(* IEC 61131-3 sources: veristc/veri-stc/tests/st-examples (part 3) *)

cond_a := LimitHigh(raw_070_a, 130);
cond_a := cond_a AND quality_a;
cond_a := cond_a AND (NOT bypass_a);
input_valid_a := InputValid(raw_070_a, 0, 1000);
cond_a := cond_a AND input_valid_a;
IF NOT input_valid_a THEN
    channel_fault_a := channel_fault_a + 1;
END_IF;
cond_b := LimitHigh(raw_070_b, 130);
cond_b := cond_b AND quality_b;
cond_b := cond_b AND (NOT bypass_b);
input_valid_b := InputValid(raw_070_b, 0, 1000);
cond_b := cond_b AND input_valid_b;
IF NOT input_valid_b THEN
    channel_fault_b := channel_fault_b + 1;
END_IF;
cond_c := LimitHigh(raw_070_c, 130);
cond_c := cond_c AND quality_c;
cond_c := cond_c AND (NOT bypass_c);
input_valid_c := InputValid(raw_070_c, 0, 1000);
cond_c := cond_c AND input_valid_c;
IF NOT input_valid_c THEN
    channel_fault_c := channel_fault_c + 1;
END_IF;
cond_d := LimitHigh(raw_070_d, 130);
cond_d := cond_d AND quality_d;
cond_d := cond_d AND (NOT bypass_d);
input_valid_d := InputValid(raw_070_d, 0, 1000);
cond_d := cond_d AND input_valid_d;
IF NOT input_valid_d THEN
    channel_fault_d := channel_fault_d + 1;
END_IF;
vote_ok := TwoOfFour(cond_a, cond_b, cond_c, cond_d);
IF cond_a <> cond_b THEN
    diagnosis_count := diagnosis_count + 1;
END_IF;
IF cond_c <> cond_d THEN
    diagnosis_count := diagnosis_count + 1;
END_IF;
IF NOT vote_ok THEN
    diagnosis_count := diagnosis_count + 1;
END_IF;
latch_a_070 := RS_Next(vote_ok, train_a_reset, latch_a_070);
IF latch_a_070 AND (NOT train_a_inhibit) THEN
    mask_a_08 := mask_a_08 + 64;
    trip_a := 0 < 1;
    scram_a := 0 < 1;
    breaker_a := 0 > 1;
    mfw_a := 0 < 1;
    alarm_a := 0 < 1;
END_IF;
latch_b_070 := RS_Next(vote_ok, train_b_reset, latch_b_070);
IF latch_b_070 AND (NOT train_b_inhibit) THEN
    mask_b_08 := mask_b_08 + 64;
    trip_b := 0 < 1;
    scram_b := 0 < 1;
    breaker_b := 0 > 1;
    mfw_b := 0 < 1;
    alarm_b := 0 < 1;
END_IF;
IF (raw_070_a > 130) AND (NOT cond_a) THEN
    channel_fault_a := channel_fault_a + 1;
END_IF;
IF (raw_070_b > 130) AND (NOT cond_b) THEN
    channel_fault_b := channel_fault_b + 1;
END_IF;
IF (raw_070_c > 130) AND (NOT cond_c) THEN
    channel_fault_c := channel_fault_c + 1;
END_IF;
IF (raw_070_d > 130) AND (NOT cond_d) THEN
    channel_fault_d := channel_fault_d + 1;
END_IF;
IF vote_ok AND train_a_inhibit THEN
    diagnosis_count := diagnosis_count + 1;
END_IF;
IF vote_ok AND train_b_inhibit THEN
    diagnosis_count := diagnosis_count + 1;
END_IF;

cond_a := LimitHigh(raw_071_a, 131);
cond_a := cond_a AND quality_a;
cond_a := cond_a AND (NOT bypass_a);
input_valid_a := InputValid(raw_071_a, 0, 1000);
cond_a := cond_a AND input_valid_a;
IF NOT input_valid_a THEN
    channel_fault_a := channel_fault_a + 1;
END_IF;
cond_b := LimitHigh(raw_071_b, 131);
cond_b := cond_b AND quality_b;
cond_b := cond_b AND (NOT bypass_b);
input_valid_b := InputValid(raw_071_b, 0, 1000);
cond_b := cond_b AND input_valid_b;
IF NOT input_valid_b THEN
    channel_fault_b := channel_fault_b + 1;
END_IF;
cond_c := LimitHigh(raw_071_c, 131);
cond_c := cond_c AND quality_c;
cond_c := cond_c AND (NOT bypass_c);
input_valid_c := InputValid(raw_071_c, 0, 1000);
cond_c := cond_c AND input_valid_c;
IF NOT input_valid_c THEN
    channel_fault_c := channel_fault_c + 1;
END_IF;
cond_d := LimitHigh(raw_071_d, 131);
cond_d := cond_d AND quality_d;
cond_d := cond_d AND (NOT bypass_d);
input_valid_d := InputValid(raw_071_d, 0, 1000);
cond_d := cond_d AND input_valid_d;
IF NOT input_valid_d THEN
    channel_fault_d := channel_fault_d + 1;
END_IF;
vote_ok := TwoOfFour(cond_a, cond_b, cond_c, cond_d);
IF cond_a <> cond_b THEN
    diagnosis_count := diagnosis_count + 1;
END_IF;
IF cond_c <> cond_d THEN
    diagnosis_count := diagnosis_count + 1;
END_IF;
IF NOT vote_ok THEN
    diagnosis_count := diagnosis_count + 1;
END_IF;
latch_a_071 := RS_Next(vote_ok, train_a_reset, latch_a_071);
IF latch_a_071 AND (NOT train_a_inhibit) THEN
    mask_a_08 := mask_a_08 + 128;
    trip_a := 0 < 1;
    scram_a := 0 < 1;
    breaker_a := 0 > 1;
    afw_a := 0 < 1;
    alarm_a := 0 < 1;
END_IF;
latch_b_071 := RS_Next(vote_ok, train_b_reset, latch_b_071);
IF latch_b_071 AND (NOT train_b_inhibit) THEN
    mask_b_08 := mask_b_08 + 128;
    trip_b := 0 < 1;
    scram_b := 0 < 1;
    breaker_b := 0 > 1;
    afw_b := 0 < 1;
    alarm_b := 0 < 1;
END_IF;
IF (raw_071_a > 131) AND (NOT cond_a) THEN
    channel_fault_a := channel_fault_a + 1;
END_IF;
IF (raw_071_b > 131) AND (NOT cond_b) THEN
    channel_fault_b := channel_fault_b + 1;
END_IF;
IF (raw_071_c > 131) AND (NOT cond_c) THEN
    channel_fault_c := channel_fault_c + 1;
END_IF;
IF (raw_071_d > 131) AND (NOT cond_d) THEN
    channel_fault_d := channel_fault_d + 1;
END_IF;
IF vote_ok AND train_a_inhibit THEN
    diagnosis_count := diagnosis_count + 1;
END_IF;
IF vote_ok AND train_b_inhibit THEN
    diagnosis_count := diagnosis_count + 1;
END_IF;

cond_a := LimitHigh(raw_072_a, 132);
cond_a := cond_a AND quality_a;
cond_a := cond_a AND (NOT bypass_a);
input_valid_a := InputValid(raw_072_a, 0, 1000);
cond_a := cond_a AND input_valid_a;
IF NOT input_valid_a THEN
    channel_fault_a := channel_fault_a + 1;
END_IF;
cond_b := LimitHigh(raw_072_b, 132);
cond_b := cond_b AND quality_b;
cond_b := cond_b AND (NOT bypass_b);
input_valid_b := InputValid(raw_072_b, 0, 1000);
cond_b := cond_b AND input_valid_b;
IF NOT input_valid_b THEN
    channel_fault_b := channel_fault_b + 1;
END_IF;
cond_c := LimitHigh(raw_072_c, 132);
cond_c := cond_c AND quality_c;
cond_c := cond_c AND (NOT bypass_c);
input_valid_c := InputValid(raw_072_c, 0, 1000);
cond_c := cond_c AND input_valid_c;
IF NOT input_valid_c THEN
    channel_fault_c := channel_fault_c + 1;
END_IF;
cond_d := LimitHigh(raw_072_d, 132);
cond_d := cond_d AND quality_d;
cond_d := cond_d AND (NOT bypass_d);
input_valid_d := InputValid(raw_072_d, 0, 1000);
cond_d := cond_d AND input_valid_d;
IF NOT input_valid_d THEN
    channel_fault_d := channel_fault_d + 1;
END_IF;
vote_ok := TwoOfFour(cond_a, cond_b, cond_c, cond_d);
IF cond_a <> cond_b THEN
    diagnosis_count := diagnosis_count + 1;
END_IF;
IF cond_c <> cond_d THEN
    diagnosis_count := diagnosis_count + 1;
END_IF;
IF NOT vote_ok THEN
    diagnosis_count := diagnosis_count + 1;
END_IF;
latch_a_072 := RS_Next(vote_ok, train_a_reset, latch_a_072);
IF latch_a_072 AND (NOT train_a_inhibit) THEN
    mask_a_09 := mask_a_09 + 1;
    trip_a := 0 < 1;
    scram_a := 0 < 1;
    breaker_a := 0 > 1;
    si_a := 0 < 1;
    alarm_a := 0 < 1;
END_IF;
latch_b_072 := RS_Next(vote_ok, train_b_reset, latch_b_072);
IF latch_b_072 AND (NOT train_b_inhibit) THEN
    mask_b_09 := mask_b_09 + 1;
    trip_b := 0 < 1;
    scram_b := 0 < 1;
    breaker_b := 0 > 1;
    si_b := 0 < 1;
    alarm_b := 0 < 1;
END_IF;
IF (raw_072_a > 132) AND (NOT cond_a) THEN
    channel_fault_a := channel_fault_a + 1;
END_IF;
IF (raw_072_b > 132) AND (NOT cond_b) THEN
    channel_fault_b := channel_fault_b + 1;
END_IF;
IF (raw_072_c > 132) AND (NOT cond_c) THEN
    channel_fault_c := channel_fault_c + 1;
END_IF;
IF (raw_072_d > 132) AND (NOT cond_d) THEN
    channel_fault_d := channel_fault_d + 1;
END_IF;
IF vote_ok AND train_a_inhibit THEN
    diagnosis_count := diagnosis_count + 1;
END_IF;
IF vote_ok AND train_b_inhibit THEN
    diagnosis_count := diagnosis_count + 1;
END_IF;

cond_a := LimitHigh(raw_073_a, 133);
cond_a := cond_a AND quality_a;
cond_a := cond_a AND (NOT bypass_a);
input_valid_a := InputValid(raw_073_a, 0, 1000);
cond_a := cond_a AND input_valid_a;
IF NOT input_valid_a THEN
    channel_fault_a := channel_fault_a + 1;
END_IF;
cond_b := LimitHigh(raw_073_b, 133);
cond_b := cond_b AND quality_b;
cond_b := cond_b AND (NOT bypass_b);
input_valid_b := InputValid(raw_073_b, 0, 1000);
cond_b := cond_b AND input_valid_b;
IF NOT input_valid_b THEN
    channel_fault_b := channel_fault_b + 1;
END_IF;
cond_c := LimitHigh(raw_073_c, 133);
cond_c := cond_c AND quality_c;
cond_c := cond_c AND (NOT bypass_c);
input_valid_c := InputValid(raw_073_c, 0, 1000);
cond_c := cond_c AND input_valid_c;
IF NOT input_valid_c THEN
    channel_fault_c := channel_fault_c + 1;
END_IF;
cond_d := LimitHigh(raw_073_d, 133);
cond_d := cond_d AND quality_d;
cond_d := cond_d AND (NOT bypass_d);
input_valid_d := InputValid(raw_073_d, 0, 1000);
cond_d := cond_d AND input_valid_d;
IF NOT input_valid_d THEN
    channel_fault_d := channel_fault_d + 1;
END_IF;
vote_ok := TwoOfFour(cond_a, cond_b, cond_c, cond_d);
IF cond_a <> cond_b THEN
    diagnosis_count := diagnosis_count + 1;
END_IF;
IF cond_c <> cond_d THEN
    diagnosis_count := diagnosis_count + 1;
END_IF;
IF NOT vote_ok THEN
    diagnosis_count := diagnosis_count + 1;
END_IF;
latch_a_073 := RS_Next(vote_ok, train_a_reset, latch_a_073);
IF latch_a_073 AND (NOT train_a_inhibit) THEN
    mask_a_09 := mask_a_09 + 2;
    trip_a := 0 < 1;
    scram_a := 0 < 1;
    breaker_a := 0 > 1;
    ci_a := 0 < 1;
    alarm_a := 0 < 1;
END_IF;
latch_b_073 := RS_Next(vote_ok, train_b_reset, latch_b_073);
IF latch_b_073 AND (NOT train_b_inhibit) THEN
    mask_b_09 := mask_b_09 + 2;
    trip_b := 0 < 1;
    scram_b := 0 < 1;
    breaker_b := 0 > 1;
    ci_b := 0 < 1;
    alarm_b := 0 < 1;
END_IF;
IF (raw_073_a > 133) AND (NOT cond_a) THEN
    channel_fault_a := channel_fault_a + 1;
END_IF;
IF (raw_073_b > 133) AND (NOT cond_b) THEN
    channel_fault_b := channel_fault_b + 1;
END_IF;
IF (raw_073_c > 133) AND (NOT cond_c) THEN
    channel_fault_c := channel_fault_c + 1;
END_IF;
IF (raw_073_d > 133) AND (NOT cond_d) THEN
    channel_fault_d := channel_fault_d + 1;
END_IF;
IF vote_ok AND train_a_inhibit THEN
    diagnosis_count := diagnosis_count + 1;
END_IF;
IF vote_ok AND train_b_inhibit THEN
    diagnosis_count := diagnosis_count + 1;
END_IF;

cond_a := LimitHigh(raw_074_a, 134);
cond_a := cond_a AND quality_a;
cond_a := cond_a AND (NOT bypass_a);
input_valid_a := InputValid(raw_074_a, 0, 1000);
cond_a := cond_a AND input_valid_a;
IF NOT input_valid_a THEN
    channel_fault_a := channel_fault_a + 1;
END_IF;
cond_b := LimitHigh(raw_074_b, 134);
cond_b := cond_b AND quality_b;
cond_b := cond_b AND (NOT bypass_b);
input_valid_b := InputValid(raw_074_b, 0, 1000);
cond_b := cond_b AND input_valid_b;
IF NOT input_valid_b THEN
    channel_fault_b := channel_fault_b + 1;
END_IF;
cond_c := LimitHigh(raw_074_c, 134);
cond_c := cond_c AND quality_c;
cond_c := cond_c AND (NOT bypass_c);
input_valid_c := InputValid(raw_074_c, 0, 1000);
cond_c := cond_c AND input_valid_c;
IF NOT input_valid_c THEN
    channel_fault_c := channel_fault_c + 1;
END_IF;
cond_d := LimitHigh(raw_074_d, 134);
cond_d := cond_d AND quality_d;
cond_d := cond_d AND (NOT bypass_d);
input_valid_d := InputValid(raw_074_d, 0, 1000);
cond_d := cond_d AND input_valid_d;
IF NOT input_valid_d THEN
    channel_fault_d := channel_fault_d + 1;
END_IF;
vote_ok := TwoOfFour(cond_a, cond_b, cond_c, cond_d);
IF cond_a <> cond_b THEN
    diagnosis_count := diagnosis_count + 1;
END_IF;
IF cond_c <> cond_d THEN
    diagnosis_count := diagnosis_count + 1;
END_IF;
IF NOT vote_ok THEN
    diagnosis_count := diagnosis_count + 1;
END_IF;
latch_a_074 := RS_Next(vote_ok, train_a_reset, latch_a_074);
IF latch_a_074 AND (NOT train_a_inhibit) THEN
    mask_a_09 := mask_a_09 + 4;
    trip_a := 0 < 1;
    scram_a := 0 < 1;
    breaker_a := 0 > 1;
    mfw_a := 0 < 1;
    alarm_a := 0 < 1;
END_IF;
latch_b_074 := RS_Next(vote_ok, train_b_reset, latch_b_074);
IF latch_b_074 AND (NOT train_b_inhibit) THEN
    mask_b_09 := mask_b_09 + 4;
    trip_b := 0 < 1;
    scram_b := 0 < 1;
    breaker_b := 0 > 1;
    mfw_b := 0 < 1;
    alarm_b := 0 < 1;
END_IF;
IF (raw_074_a > 134) AND (NOT cond_a) THEN
    channel_fault_a := channel_fault_a + 1;
END_IF;
IF (raw_074_b > 134) AND (NOT cond_b) THEN
    channel_fault_b := channel_fault_b + 1;
END_IF;
IF (raw_074_c > 134) AND (NOT cond_c) THEN
    channel_fault_c := channel_fault_c + 1;
END_IF;
IF (raw_074_d > 134) AND (NOT cond_d) THEN
    channel_fault_d := channel_fault_d + 1;
END_IF;
IF vote_ok AND train_a_inhibit THEN
    diagnosis_count := diagnosis_count + 1;
END_IF;
IF vote_ok AND train_b_inhibit THEN
    diagnosis_count := diagnosis_count + 1;
END_IF;

cond_a := LimitHigh(raw_075_a, 135);
cond_a := cond_a AND quality_a;
cond_a := cond_a AND (NOT bypass_a);
input_valid_a := InputValid(raw_075_a, 0, 1000);
cond_a := cond_a AND input_valid_a;
IF NOT input_valid_a THEN
    channel_fault_a := channel_fault_a + 1;
END_IF;
cond_b := LimitHigh(raw_075_b, 135);
cond_b := cond_b AND quality_b;
cond_b := cond_b AND (NOT bypass_b);
input_valid_b := InputValid(raw_075_b, 0, 1000);
cond_b := cond_b AND input_valid_b;
IF NOT input_valid_b THEN
    channel_fault_b := channel_fault_b + 1;
END_IF;
cond_c := LimitHigh(raw_075_c, 135);
cond_c := cond_c AND quality_c;
cond_c := cond_c AND (NOT bypass_c);
input_valid_c := InputValid(raw_075_c, 0, 1000);
cond_c := cond_c AND input_valid_c;
IF NOT input_valid_c THEN
    channel_fault_c := channel_fault_c + 1;
END_IF;
cond_d := LimitHigh(raw_075_d, 135);
cond_d := cond_d AND quality_d;
cond_d := cond_d AND (NOT bypass_d);
input_valid_d := InputValid(raw_075_d, 0, 1000);
cond_d := cond_d AND input_valid_d;
IF NOT input_valid_d THEN
    channel_fault_d := channel_fault_d + 1;
END_IF;
vote_ok := TwoOfFour(cond_a, cond_b, cond_c, cond_d);
IF cond_a <> cond_b THEN
    diagnosis_count := diagnosis_count + 1;
END_IF;
IF cond_c <> cond_d THEN
    diagnosis_count := diagnosis_count + 1;
END_IF;
IF NOT vote_ok THEN
    diagnosis_count := diagnosis_count + 1;
END_IF;
latch_a_075 := RS_Next(vote_ok, train_a_reset, latch_a_075);
IF latch_a_075 AND (NOT train_a_inhibit) THEN
    mask_a_09 := mask_a_09 + 8;
    trip_a := 0 < 1;
    scram_a := 0 < 1;
    breaker_a := 0 > 1;
    afw_a := 0 < 1;
    alarm_a := 0 < 1;
END_IF;
latch_b_075 := RS_Next(vote_ok, train_b_reset, latch_b_075);
IF latch_b_075 AND (NOT train_b_inhibit) THEN
    mask_b_09 := mask_b_09 + 8;
    trip_b := 0 < 1;
    scram_b := 0 < 1;
    breaker_b := 0 > 1;
    afw_b := 0 < 1;
    alarm_b := 0 < 1;
END_IF;
IF (raw_075_a > 135) AND (NOT cond_a) THEN
    channel_fault_a := channel_fault_a + 1;
END_IF;
IF (raw_075_b > 135) AND (NOT cond_b) THEN
    channel_fault_b := channel_fault_b + 1;
END_IF;
IF (raw_075_c > 135) AND (NOT cond_c) THEN
    channel_fault_c := channel_fault_c + 1;
END_IF;
IF (raw_075_d > 135) AND (NOT cond_d) THEN
    channel_fault_d := channel_fault_d + 1;
END_IF;
IF vote_ok AND train_a_inhibit THEN
    diagnosis_count := diagnosis_count + 1;
END_IF;
IF vote_ok AND train_b_inhibit THEN
    diagnosis_count := diagnosis_count + 1;
END_IF;

cond_a := LimitHigh(raw_076_a, 136);
cond_a := cond_a AND quality_a;
cond_a := cond_a AND (NOT bypass_a);
input_valid_a := InputValid(raw_076_a, 0, 1000);
cond_a := cond_a AND input_valid_a;
IF NOT input_valid_a THEN
    channel_fault_a := channel_fault_a + 1;
END_IF;
cond_b := LimitHigh(raw_076_b, 136);
cond_b := cond_b AND quality_b;
cond_b := cond_b AND (NOT bypass_b);
input_valid_b := InputValid(raw_076_b, 0, 1000);
cond_b := cond_b AND input_valid_b;
IF NOT input_valid_b THEN
    channel_fault_b := channel_fault_b + 1;
END_IF;
cond_c := LimitHigh(raw_076_c, 136);
cond_c := cond_c AND quality_c;
cond_c := cond_c AND (NOT bypass_c);
input_valid_c := InputValid(raw_076_c, 0, 1000);
cond_c := cond_c AND input_valid_c;
IF NOT input_valid_c THEN
    channel_fault_c := channel_fault_c + 1;
END_IF;
cond_d := LimitHigh(raw_076_d, 136);
cond_d := cond_d AND quality_d;
cond_d := cond_d AND (NOT bypass_d);
input_valid_d := InputValid(raw_076_d, 0, 1000);
cond_d := cond_d AND input_valid_d;
IF NOT input_valid_d THEN
    channel_fault_d := channel_fault_d + 1;
END_IF;
vote_ok := TwoOfFour(cond_a, cond_b, cond_c, cond_d);
IF cond_a <> cond_b THEN
    diagnosis_count := diagnosis_count + 1;
END_IF;
IF cond_c <> cond_d THEN
    diagnosis_count := diagnosis_count + 1;
END_IF;
IF NOT vote_ok THEN
    diagnosis_count := diagnosis_count + 1;
END_IF;
latch_a_076 := RS_Next(vote_ok, train_a_reset, latch_a_076);
IF latch_a_076 AND (NOT train_a_inhibit) THEN
    mask_a_09 := mask_a_09 + 16;
    trip_a := 0 < 1;
    scram_a := 0 < 1;
    breaker_a := 0 > 1;
    si_a := 0 < 1;
    alarm_a := 0 < 1;
END_IF;
latch_b_076 := RS_Next(vote_ok, train_b_reset, latch_b_076);
IF latch_b_076 AND (NOT train_b_inhibit) THEN
    mask_b_09 := mask_b_09 + 16;
    trip_b := 0 < 1;
    scram_b := 0 < 1;
    breaker_b := 0 > 1;
    si_b := 0 < 1;
    alarm_b := 0 < 1;
END_IF;
IF (raw_076_a > 136) AND (NOT cond_a) THEN
    channel_fault_a := channel_fault_a + 1;
END_IF;
IF (raw_076_b > 136) AND (NOT cond_b) THEN
    channel_fault_b := channel_fault_b + 1;
END_IF;
IF (raw_076_c > 136) AND (NOT cond_c) THEN
    channel_fault_c := channel_fault_c + 1;
END_IF;
IF (raw_076_d > 136) AND (NOT cond_d) THEN
    channel_fault_d := channel_fault_d + 1;
END_IF;
IF vote_ok AND train_a_inhibit THEN
    diagnosis_count := diagnosis_count + 1;
END_IF;
IF vote_ok AND train_b_inhibit THEN
    diagnosis_count := diagnosis_count + 1;
END_IF;

cond_a := LimitHigh(raw_077_a, 137);
cond_a := cond_a AND quality_a;
cond_a := cond_a AND (NOT bypass_a);
input_valid_a := InputValid(raw_077_a, 0, 1000);
cond_a := cond_a AND input_valid_a;
IF NOT input_valid_a THEN
    channel_fault_a := channel_fault_a + 1;
END_IF;
cond_b := LimitHigh(raw_077_b, 137);
cond_b := cond_b AND quality_b;
cond_b := cond_b AND (NOT bypass_b);
input_valid_b := InputValid(raw_077_b, 0, 1000);
cond_b := cond_b AND input_valid_b;
IF NOT input_valid_b THEN
    channel_fault_b := channel_fault_b + 1;
END_IF;
cond_c := LimitHigh(raw_077_c, 137);
cond_c := cond_c AND quality_c;
cond_c := cond_c AND (NOT bypass_c);
input_valid_c := InputValid(raw_077_c, 0, 1000);
cond_c := cond_c AND input_valid_c;
IF NOT input_valid_c THEN
    channel_fault_c := channel_fault_c + 1;
END_IF;
cond_d := LimitHigh(raw_077_d, 137);
cond_d := cond_d AND quality_d;
cond_d := cond_d AND (NOT bypass_d);
input_valid_d := InputValid(raw_077_d, 0, 1000);
cond_d := cond_d AND input_valid_d;
IF NOT input_valid_d THEN
    channel_fault_d := channel_fault_d + 1;
END_IF;
vote_ok := TwoOfFour(cond_a, cond_b, cond_c, cond_d);
IF cond_a <> cond_b THEN
    diagnosis_count := diagnosis_count + 1;
END_IF;
IF cond_c <> cond_d THEN
    diagnosis_count := diagnosis_count + 1;
END_IF;
IF NOT vote_ok THEN
    diagnosis_count := diagnosis_count + 1;
END_IF;
latch_a_077 := RS_Next(vote_ok, train_a_reset, latch_a_077);
IF latch_a_077 AND (NOT train_a_inhibit) THEN
    mask_a_09 := mask_a_09 + 32;
    trip_a := 0 < 1;
    scram_a := 0 < 1;
    breaker_a := 0 > 1;
    ci_a := 0 < 1;
    alarm_a := 0 < 1;
END_IF;
latch_b_077 := RS_Next(vote_ok, train_b_reset, latch_b_077);
IF latch_b_077 AND (NOT train_b_inhibit) THEN
    mask_b_09 := mask_b_09 + 32;
    trip_b := 0 < 1;
    scram_b := 0 < 1;
    breaker_b := 0 > 1;
    ci_b := 0 < 1;
    alarm_b := 0 < 1;
END_IF;
IF (raw_077_a > 137) AND (NOT cond_a) THEN
    channel_fault_a := channel_fault_a + 1;
END_IF;
IF (raw_077_b > 137) AND (NOT cond_b) THEN
    channel_fault_b := channel_fault_b + 1;
END_IF;
IF (raw_077_c > 137) AND (NOT cond_c) THEN
    channel_fault_c := channel_fault_c + 1;
END_IF;
IF (raw_077_d > 137) AND (NOT cond_d) THEN
    channel_fault_d := channel_fault_d + 1;
END_IF;
IF vote_ok AND train_a_inhibit THEN
    diagnosis_count := diagnosis_count + 1;
END_IF;
IF vote_ok AND train_b_inhibit THEN
    diagnosis_count := diagnosis_count + 1;
END_IF;

cond_a := LimitHigh(raw_078_a, 138);
cond_a := cond_a AND quality_a;
cond_a := cond_a AND (NOT bypass_a);
input_valid_a := InputValid(raw_078_a, 0, 1000);
cond_a := cond_a AND input_valid_a;
IF NOT input_valid_a THEN
    channel_fault_a := channel_fault_a + 1;
END_IF;
cond_b := LimitHigh(raw_078_b, 138);
cond_b := cond_b AND quality_b;
cond_b := cond_b AND (NOT bypass_b);
input_valid_b := InputValid(raw_078_b, 0, 1000);
cond_b := cond_b AND input_valid_b;
IF NOT input_valid_b THEN
    channel_fault_b := channel_fault_b + 1;
END_IF;
cond_c := LimitHigh(raw_078_c, 138);
cond_c := cond_c AND quality_c;
cond_c := cond_c AND (NOT bypass_c);
input_valid_c := InputValid(raw_078_c, 0, 1000);
cond_c := cond_c AND input_valid_c;
IF NOT input_valid_c THEN
    channel_fault_c := channel_fault_c + 1;
END_IF;
cond_d := LimitHigh(raw_078_d, 138);
cond_d := cond_d AND quality_d;
cond_d := cond_d AND (NOT bypass_d);
input_valid_d := InputValid(raw_078_d, 0, 1000);
cond_d := cond_d AND input_valid_d;
IF NOT input_valid_d THEN
    channel_fault_d := channel_fault_d + 1;
END_IF;
vote_ok := TwoOfFour(cond_a, cond_b, cond_c, cond_d);
IF cond_a <> cond_b THEN
    diagnosis_count := diagnosis_count + 1;
END_IF;
IF cond_c <> cond_d THEN
    diagnosis_count := diagnosis_count + 1;
END_IF;
IF NOT vote_ok THEN
    diagnosis_count := diagnosis_count + 1;
END_IF;
latch_a_078 := RS_Next(vote_ok, train_a_reset, latch_a_078);
IF latch_a_078 AND (NOT train_a_inhibit) THEN
    mask_a_09 := mask_a_09 + 64;
    trip_a := 0 < 1;
    scram_a := 0 < 1;
    breaker_a := 0 > 1;
    mfw_a := 0 < 1;
    alarm_a := 0 < 1;
END_IF;
latch_b_078 := RS_Next(vote_ok, train_b_reset, latch_b_078);
IF latch_b_078 AND (NOT train_b_inhibit) THEN
    mask_b_09 := mask_b_09 + 64;
    trip_b := 0 < 1;
    scram_b := 0 < 1;
    breaker_b := 0 > 1;
    mfw_b := 0 < 1;
    alarm_b := 0 < 1;
END_IF;
IF (raw_078_a > 138) AND (NOT cond_a) THEN
    channel_fault_a := channel_fault_a + 1;
END_IF;
IF (raw_078_b > 138) AND (NOT cond_b) THEN
    channel_fault_b := channel_fault_b + 1;
END_IF;
IF (raw_078_c > 138) AND (NOT cond_c) THEN
    channel_fault_c := channel_fault_c + 1;
END_IF;
IF (raw_078_d > 138) AND (NOT cond_d) THEN
    channel_fault_d := channel_fault_d + 1;
END_IF;
IF vote_ok AND train_a_inhibit THEN
    diagnosis_count := diagnosis_count + 1;
END_IF;
IF vote_ok AND train_b_inhibit THEN
    diagnosis_count := diagnosis_count + 1;
END_IF;

cond_a := LimitHigh(raw_079_a, 139);
cond_a := cond_a AND quality_a;
cond_a := cond_a AND (NOT bypass_a);
input_valid_a := InputValid(raw_079_a, 0, 1000);
cond_a := cond_a AND input_valid_a;
IF NOT input_valid_a THEN
    channel_fault_a := channel_fault_a + 1;
END_IF;
cond_b := LimitHigh(raw_079_b, 139);
cond_b := cond_b AND quality_b;
cond_b := cond_b AND (NOT bypass_b);
input_valid_b := InputValid(raw_079_b, 0, 1000);
cond_b := cond_b AND input_valid_b;
IF NOT input_valid_b THEN
    channel_fault_b := channel_fault_b + 1;
END_IF;
cond_c := LimitHigh(raw_079_c, 139);
cond_c := cond_c AND quality_c;
cond_c := cond_c AND (NOT bypass_c);
input_valid_c := InputValid(raw_079_c, 0, 1000);
cond_c := cond_c AND input_valid_c;
IF NOT input_valid_c THEN
    channel_fault_c := channel_fault_c + 1;
END_IF;
cond_d := LimitHigh(raw_079_d, 139);
cond_d := cond_d AND quality_d;
cond_d := cond_d AND (NOT bypass_d);
input_valid_d := InputValid(raw_079_d, 0, 1000);
cond_d := cond_d AND input_valid_d;
IF NOT input_valid_d THEN
    channel_fault_d := channel_fault_d + 1;
END_IF;
vote_ok := TwoOfFour(cond_a, cond_b, cond_c, cond_d);
IF cond_a <> cond_b THEN
    diagnosis_count := diagnosis_count + 1;
END_IF;
IF cond_c <> cond_d THEN
    diagnosis_count := diagnosis_count + 1;
END_IF;
IF NOT vote_ok THEN
    diagnosis_count := diagnosis_count + 1;
END_IF;
latch_a_079 := RS_Next(vote_ok, train_a_reset, latch_a_079);
IF latch_a_079 AND (NOT train_a_inhibit) THEN
    mask_a_09 := mask_a_09 + 128;
    trip_a := 0 < 1;
    scram_a := 0 < 1;
    breaker_a := 0 > 1;
    afw_a := 0 < 1;
    alarm_a := 0 < 1;
END_IF;
latch_b_079 := RS_Next(vote_ok, train_b_reset, latch_b_079);
IF latch_b_079 AND (NOT train_b_inhibit) THEN
    mask_b_09 := mask_b_09 + 128;
    trip_b := 0 < 1;
    scram_b := 0 < 1;
    breaker_b := 0 > 1;
    afw_b := 0 < 1;
    alarm_b := 0 < 1;
END_IF;
IF (raw_079_a > 139) AND (NOT cond_a) THEN
    channel_fault_a := channel_fault_a + 1;
END_IF;
IF (raw_079_b > 139) AND (NOT cond_b) THEN
    channel_fault_b := channel_fault_b + 1;
END_IF;
IF (raw_079_c > 139) AND (NOT cond_c) THEN
    channel_fault_c := channel_fault_c + 1;
END_IF;
IF (raw_079_d > 139) AND (NOT cond_d) THEN
    channel_fault_d := channel_fault_d + 1;
END_IF;
IF vote_ok AND train_a_inhibit THEN
    diagnosis_count := diagnosis_count + 1;
END_IF;
IF vote_ok AND train_b_inhibit THEN
    diagnosis_count := diagnosis_count + 1;
END_IF;

cond_a := LimitHigh(raw_080_a, 100);
cond_a := cond_a AND quality_a;
cond_a := cond_a AND (NOT bypass_a);
input_valid_a := InputValid(raw_080_a, 0, 1000);
cond_a := cond_a AND input_valid_a;
IF NOT input_valid_a THEN
    channel_fault_a := channel_fault_a + 1;
END_IF;
cond_b := LimitHigh(raw_080_b, 100);
cond_b := cond_b AND quality_b;
cond_b := cond_b AND (NOT bypass_b);
input_valid_b := InputValid(raw_080_b, 0, 1000);
cond_b := cond_b AND input_valid_b;
IF NOT input_valid_b THEN
    channel_fault_b := channel_fault_b + 1;
END_IF;
cond_c := LimitHigh(raw_080_c, 100);
cond_c := cond_c AND quality_c;
cond_c := cond_c AND (NOT bypass_c);
input_valid_c := InputValid(raw_080_c, 0, 1000);
cond_c := cond_c AND input_valid_c;
IF NOT input_valid_c THEN
    channel_fault_c := channel_fault_c + 1;
END_IF;
cond_d := LimitHigh(raw_080_d, 100);
cond_d := cond_d AND quality_d;
cond_d := cond_d AND (NOT bypass_d);
input_valid_d := InputValid(raw_080_d, 0, 1000);
cond_d := cond_d AND input_valid_d;
IF NOT input_valid_d THEN
    channel_fault_d := channel_fault_d + 1;
END_IF;
vote_ok := TwoOfFour(cond_a, cond_b, cond_c, cond_d);
IF cond_a <> cond_b THEN
    diagnosis_count := diagnosis_count + 1;
END_IF;
IF cond_c <> cond_d THEN
    diagnosis_count := diagnosis_count + 1;
END_IF;
IF NOT vote_ok THEN
    diagnosis_count := diagnosis_count + 1;
END_IF;
latch_a_080 := RS_Next(vote_ok, train_a_reset, latch_a_080);
IF latch_a_080 AND (NOT train_a_inhibit) THEN
    mask_a_10 := mask_a_10 + 1;
    trip_a := 0 < 1;
    scram_a := 0 < 1;
    breaker_a := 0 > 1;
    si_a := 0 < 1;
    alarm_a := 0 < 1;
END_IF;
latch_b_080 := RS_Next(vote_ok, train_b_reset, latch_b_080);
IF latch_b_080 AND (NOT train_b_inhibit) THEN
    mask_b_10 := mask_b_10 + 1;
    trip_b := 0 < 1;
    scram_b := 0 < 1;
    breaker_b := 0 > 1;
    si_b := 0 < 1;
    alarm_b := 0 < 1;
END_IF;
IF (raw_080_a > 100) AND (NOT cond_a) THEN
    channel_fault_a := channel_fault_a + 1;
END_IF;
IF (raw_080_b > 100) AND (NOT cond_b) THEN
    channel_fault_b := channel_fault_b + 1;
END_IF;
IF (raw_080_c > 100) AND (NOT cond_c) THEN
    channel_fault_c := channel_fault_c + 1;
END_IF;
IF (raw_080_d > 100) AND (NOT cond_d) THEN
    channel_fault_d := channel_fault_d + 1;
END_IF;
IF vote_ok AND train_a_inhibit THEN
    diagnosis_count := diagnosis_count + 1;
END_IF;
IF vote_ok AND train_b_inhibit THEN
    diagnosis_count := diagnosis_count + 1;
END_IF;

cond_a := LimitHigh(raw_081_a, 101);
cond_a := cond_a AND quality_a;
cond_a := cond_a AND (NOT bypass_a);
input_valid_a := InputValid(raw_081_a, 0, 1000);
cond_a := cond_a AND input_valid_a;
IF NOT input_valid_a THEN
    channel_fault_a := channel_fault_a + 1;
END_IF;
cond_b := LimitHigh(raw_081_b, 101);
cond_b := cond_b AND quality_b;
cond_b := cond_b AND (NOT bypass_b);
input_valid_b := InputValid(raw_081_b, 0, 1000);
cond_b := cond_b AND input_valid_b;
IF NOT input_valid_b THEN
    channel_fault_b := channel_fault_b + 1;
END_IF;
cond_c := LimitHigh(raw_081_c, 101);
cond_c := cond_c AND quality_c;
cond_c := cond_c AND (NOT bypass_c);
input_valid_c := InputValid(raw_081_c, 0, 1000);
cond_c := cond_c AND input_valid_c;
IF NOT input_valid_c THEN
    channel_fault_c := channel_fault_c + 1;
END_IF;
cond_d := LimitHigh(raw_081_d, 101);
cond_d := cond_d AND quality_d;
cond_d := cond_d AND (NOT bypass_d);
input_valid_d := InputValid(raw_081_d, 0, 1000);
cond_d := cond_d AND input_valid_d;
IF NOT input_valid_d THEN
    channel_fault_d := channel_fault_d + 1;
END_IF;
vote_ok := TwoOfFour(cond_a, cond_b, cond_c, cond_d);
IF cond_a <> cond_b THEN
    diagnosis_count := diagnosis_count + 1;
END_IF;
IF cond_c <> cond_d THEN
    diagnosis_count := diagnosis_count + 1;
END_IF;
IF NOT vote_ok THEN
    diagnosis_count := diagnosis_count + 1;
END_IF;
latch_a_081 := RS_Next(vote_ok, train_a_reset, latch_a_081);
IF latch_a_081 AND (NOT train_a_inhibit) THEN
    mask_a_10 := mask_a_10 + 2;
    trip_a := 0 < 1;
    scram_a := 0 < 1;
    breaker_a := 0 > 1;
    ci_a := 0 < 1;
    alarm_a := 0 < 1;
END_IF;
latch_b_081 := RS_Next(vote_ok, train_b_reset, latch_b_081);
IF latch_b_081 AND (NOT train_b_inhibit) THEN
    mask_b_10 := mask_b_10 + 2;
    trip_b := 0 < 1;
    scram_b := 0 < 1;
    breaker_b := 0 > 1;
    ci_b := 0 < 1;
    alarm_b := 0 < 1;
END_IF;
IF (raw_081_a > 101) AND (NOT cond_a) THEN
    channel_fault_a := channel_fault_a + 1;
END_IF;
IF (raw_081_b > 101) AND (NOT cond_b) THEN
    channel_fault_b := channel_fault_b + 1;
END_IF;
IF (raw_081_c > 101) AND (NOT cond_c) THEN
    channel_fault_c := channel_fault_c + 1;
END_IF;
IF (raw_081_d > 101) AND (NOT cond_d) THEN
    channel_fault_d := channel_fault_d + 1;
END_IF;
IF vote_ok AND train_a_inhibit THEN
    diagnosis_count := diagnosis_count + 1;
END_IF;
IF vote_ok AND train_b_inhibit THEN
    diagnosis_count := diagnosis_count + 1;
END_IF;

cond_a := LimitHigh(raw_082_a, 102);
cond_a := cond_a AND quality_a;
cond_a := cond_a AND (NOT bypass_a);
input_valid_a := InputValid(raw_082_a, 0, 1000);
cond_a := cond_a AND input_valid_a;
IF NOT input_valid_a THEN
    channel_fault_a := channel_fault_a + 1;
END_IF;
cond_b := LimitHigh(raw_082_b, 102);
cond_b := cond_b AND quality_b;
cond_b := cond_b AND (NOT bypass_b);
input_valid_b := InputValid(raw_082_b, 0, 1000);
cond_b := cond_b AND input_valid_b;
IF NOT input_valid_b THEN
    channel_fault_b := channel_fault_b + 1;
END_IF;
cond_c := LimitHigh(raw_082_c, 102);
cond_c := cond_c AND quality_c;
cond_c := cond_c AND (NOT bypass_c);
input_valid_c := InputValid(raw_082_c, 0, 1000);
cond_c := cond_c AND input_valid_c;
IF NOT input_valid_c THEN
    channel_fault_c := channel_fault_c + 1;
END_IF;
cond_d := LimitHigh(raw_082_d, 102);
cond_d := cond_d AND quality_d;
cond_d := cond_d AND (NOT bypass_d);
input_valid_d := InputValid(raw_082_d, 0, 1000);
cond_d := cond_d AND input_valid_d;
IF NOT input_valid_d THEN
    channel_fault_d := channel_fault_d + 1;
END_IF;
vote_ok := TwoOfFour(cond_a, cond_b, cond_c, cond_d);
IF cond_a <> cond_b THEN
    diagnosis_count := diagnosis_count + 1;
END_IF;
IF cond_c <> cond_d THEN
    diagnosis_count := diagnosis_count + 1;
END_IF;
IF NOT vote_ok THEN
    diagnosis_count := diagnosis_count + 1;
END_IF;
latch_a_082 := RS_Next(vote_ok, train_a_reset, latch_a_082);
IF latch_a_082 AND (NOT train_a_inhibit) THEN
    mask_a_10 := mask_a_10 + 4;
    trip_a := 0 < 1;
    scram_a := 0 < 1;
    breaker_a := 0 > 1;
    mfw_a := 0 < 1;
    alarm_a := 0 < 1;
END_IF;
latch_b_082 := RS_Next(vote_ok, train_b_reset, latch_b_082);
IF latch_b_082 AND (NOT train_b_inhibit) THEN
    mask_b_10 := mask_b_10 + 4;
    trip_b := 0 < 1;
    scram_b := 0 < 1;
    breaker_b := 0 > 1;
    mfw_b := 0 < 1;
    alarm_b := 0 < 1;
END_IF;
IF (raw_082_a > 102) AND (NOT cond_a) THEN
    channel_fault_a := channel_fault_a + 1;
END_IF;
IF (raw_082_b > 102) AND (NOT cond_b) THEN
    channel_fault_b := channel_fault_b + 1;
END_IF;
IF (raw_082_c > 102) AND (NOT cond_c) THEN
    channel_fault_c := channel_fault_c + 1;
END_IF;
IF (raw_082_d > 102) AND (NOT cond_d) THEN
    channel_fault_d := channel_fault_d + 1;
END_IF;
IF vote_ok AND train_a_inhibit THEN
    diagnosis_count := diagnosis_count + 1;
END_IF;
IF vote_ok AND train_b_inhibit THEN
    diagnosis_count := diagnosis_count + 1;
END_IF;

cond_a := LimitHigh(raw_083_a, 103);
cond_a := cond_a AND quality_a;
cond_a := cond_a AND (NOT bypass_a);
input_valid_a := InputValid(raw_083_a, 0, 1000);
cond_a := cond_a AND input_valid_a;
IF NOT input_valid_a THEN
    channel_fault_a := channel_fault_a + 1;
END_IF;
cond_b := LimitHigh(raw_083_b, 103);
cond_b := cond_b AND quality_b;
cond_b := cond_b AND (NOT bypass_b);
input_valid_b := InputValid(raw_083_b, 0, 1000);
cond_b := cond_b AND input_valid_b;
IF NOT input_valid_b THEN
    channel_fault_b := channel_fault_b + 1;
END_IF;
cond_c := LimitHigh(raw_083_c, 103);
cond_c := cond_c AND quality_c;
cond_c := cond_c AND (NOT bypass_c);
input_valid_c := InputValid(raw_083_c, 0, 1000);
cond_c := cond_c AND input_valid_c;
IF NOT input_valid_c THEN
    channel_fault_c := channel_fault_c + 1;
END_IF;
cond_d := LimitHigh(raw_083_d, 103);
cond_d := cond_d AND quality_d;
cond_d := cond_d AND (NOT bypass_d);
input_valid_d := InputValid(raw_083_d, 0, 1000);
cond_d := cond_d AND input_valid_d;
IF NOT input_valid_d THEN
    channel_fault_d := channel_fault_d + 1;
END_IF;
vote_ok := TwoOfFour(cond_a, cond_b, cond_c, cond_d);
IF cond_a <> cond_b THEN
    diagnosis_count := diagnosis_count + 1;
END_IF;
IF cond_c <> cond_d THEN
    diagnosis_count := diagnosis_count + 1;
END_IF;
IF NOT vote_ok THEN
    diagnosis_count := diagnosis_count + 1;
END_IF;
latch_a_083 := RS_Next(vote_ok, train_a_reset, latch_a_083);
IF latch_a_083 AND (NOT train_a_inhibit) THEN
    mask_a_10 := mask_a_10 + 8;
    trip_a := 0 < 1;
    scram_a := 0 < 1;
    breaker_a := 0 > 1;
    afw_a := 0 < 1;
    alarm_a := 0 < 1;
END_IF;
latch_b_083 := RS_Next(vote_ok, train_b_reset, latch_b_083);
IF latch_b_083 AND (NOT train_b_inhibit) THEN
    mask_b_10 := mask_b_10 + 8;
    trip_b := 0 < 1;
    scram_b := 0 < 1;
    breaker_b := 0 > 1;
    afw_b := 0 < 1;
    alarm_b := 0 < 1;
END_IF;
IF (raw_083_a > 103) AND (NOT cond_a) THEN
    channel_fault_a := channel_fault_a + 1;
END_IF;
IF (raw_083_b > 103) AND (NOT cond_b) THEN
    channel_fault_b := channel_fault_b + 1;
END_IF;
IF (raw_083_c > 103) AND (NOT cond_c) THEN
    channel_fault_c := channel_fault_c + 1;
END_IF;
IF (raw_083_d > 103) AND (NOT cond_d) THEN
    channel_fault_d := channel_fault_d + 1;
END_IF;
IF vote_ok AND train_a_inhibit THEN
    diagnosis_count := diagnosis_count + 1;
END_IF;
IF vote_ok AND train_b_inhibit THEN
    diagnosis_count := diagnosis_count + 1;
END_IF;

cond_a := LimitHigh(raw_084_a, 104);
cond_a := cond_a AND quality_a;
cond_a := cond_a AND (NOT bypass_a);
input_valid_a := InputValid(raw_084_a, 0, 1000);
cond_a := cond_a AND input_valid_a;
IF NOT input_valid_a THEN
    channel_fault_a := channel_fault_a + 1;
END_IF;
cond_b := LimitHigh(raw_084_b, 104);
cond_b := cond_b AND quality_b;
cond_b := cond_b AND (NOT bypass_b);
input_valid_b := InputValid(raw_084_b, 0, 1000);
cond_b := cond_b AND input_valid_b;
IF NOT input_valid_b THEN
    channel_fault_b := channel_fault_b + 1;
END_IF;
cond_c := LimitHigh(raw_084_c, 104);
cond_c := cond_c AND quality_c;
cond_c := cond_c AND (NOT bypass_c);
input_valid_c := InputValid(raw_084_c, 0, 1000);
cond_c := cond_c AND input_valid_c;
IF NOT input_valid_c THEN
    channel_fault_c := channel_fault_c + 1;
END_IF;
cond_d := LimitHigh(raw_084_d, 104);
cond_d := cond_d AND quality_d;
cond_d := cond_d AND (NOT bypass_d);
input_valid_d := InputValid(raw_084_d, 0, 1000);
cond_d := cond_d AND input_valid_d;
IF NOT input_valid_d THEN
    channel_fault_d := channel_fault_d + 1;
END_IF;
vote_ok := TwoOfFour(cond_a, cond_b, cond_c, cond_d);
IF cond_a <> cond_b THEN
    diagnosis_count := diagnosis_count + 1;
END_IF;
IF cond_c <> cond_d THEN
    diagnosis_count := diagnosis_count + 1;
END_IF;
IF NOT vote_ok THEN
    diagnosis_count := diagnosis_count + 1;
END_IF;
latch_a_084 := RS_Next(vote_ok, train_a_reset, latch_a_084);
IF latch_a_084 AND (NOT train_a_inhibit) THEN
    mask_a_10 := mask_a_10 + 16;
    trip_a := 0 < 1;
    scram_a := 0 < 1;
    breaker_a := 0 > 1;
    si_a := 0 < 1;
    alarm_a := 0 < 1;
END_IF;
latch_b_084 := RS_Next(vote_ok, train_b_reset, latch_b_084);
IF latch_b_084 AND (NOT train_b_inhibit) THEN
    mask_b_10 := mask_b_10 + 16;
    trip_b := 0 < 1;
    scram_b := 0 < 1;
    breaker_b := 0 > 1;
    si_b := 0 < 1;
    alarm_b := 0 < 1;
END_IF;
IF (raw_084_a > 104) AND (NOT cond_a) THEN
    channel_fault_a := channel_fault_a + 1;
END_IF;
IF (raw_084_b > 104) AND (NOT cond_b) THEN
    channel_fault_b := channel_fault_b + 1;
END_IF;
IF (raw_084_c > 104) AND (NOT cond_c) THEN
    channel_fault_c := channel_fault_c + 1;
END_IF;
IF (raw_084_d > 104) AND (NOT cond_d) THEN
    channel_fault_d := channel_fault_d + 1;
END_IF;
IF vote_ok AND train_a_inhibit THEN
    diagnosis_count := diagnosis_count + 1;
END_IF;
IF vote_ok AND train_b_inhibit THEN
    diagnosis_count := diagnosis_count + 1;
END_IF;

cond_a := LimitHigh(raw_085_a, 105);
cond_a := cond_a AND quality_a;
cond_a := cond_a AND (NOT bypass_a);
input_valid_a := InputValid(raw_085_a, 0, 1000);
cond_a := cond_a AND input_valid_a;
IF NOT input_valid_a THEN
    channel_fault_a := channel_fault_a + 1;
END_IF;
cond_b := LimitHigh(raw_085_b, 105);
cond_b := cond_b AND quality_b;
cond_b := cond_b AND (NOT bypass_b);
input_valid_b := InputValid(raw_085_b, 0, 1000);
cond_b := cond_b AND input_valid_b;
IF NOT input_valid_b THEN
    channel_fault_b := channel_fault_b + 1;
END_IF;
cond_c := LimitHigh(raw_085_c, 105);
cond_c := cond_c AND quality_c;
cond_c := cond_c AND (NOT bypass_c);
input_valid_c := InputValid(raw_085_c, 0, 1000);
cond_c := cond_c AND input_valid_c;
IF NOT input_valid_c THEN
    channel_fault_c := channel_fault_c + 1;
END_IF;
cond_d := LimitHigh(raw_085_d, 105);
cond_d := cond_d AND quality_d;
cond_d := cond_d AND (NOT bypass_d);
input_valid_d := InputValid(raw_085_d, 0, 1000);
cond_d := cond_d AND input_valid_d;
IF NOT input_valid_d THEN
    channel_fault_d := channel_fault_d + 1;
END_IF;
vote_ok := TwoOfFour(cond_a, cond_b, cond_c, cond_d);
IF cond_a <> cond_b THEN
    diagnosis_count := diagnosis_count + 1;
END_IF;
IF cond_c <> cond_d THEN
    diagnosis_count := diagnosis_count + 1;
END_IF;
IF NOT vote_ok THEN
    diagnosis_count := diagnosis_count + 1;
END_IF;
latch_a_085 := RS_Next(vote_ok, train_a_reset, latch_a_085);
IF latch_a_085 AND (NOT train_a_inhibit) THEN
    mask_a_10 := mask_a_10 + 32;
    trip_a := 0 < 1;
    scram_a := 0 < 1;
    breaker_a := 0 > 1;
    ci_a := 0 < 1;
    alarm_a := 0 < 1;
END_IF;
latch_b_085 := RS_Next(vote_ok, train_b_reset, latch_b_085);
IF latch_b_085 AND (NOT train_b_inhibit) THEN
    mask_b_10 := mask_b_10 + 32;
    trip_b := 0 < 1;
    scram_b := 0 < 1;
    breaker_b := 0 > 1;
    ci_b := 0 < 1;
    alarm_b := 0 < 1;
END_IF;
IF (raw_085_a > 105) AND (NOT cond_a) THEN
    channel_fault_a := channel_fault_a + 1;
END_IF;
IF (raw_085_b > 105) AND (NOT cond_b) THEN
    channel_fault_b := channel_fault_b + 1;
END_IF;
IF (raw_085_c > 105) AND (NOT cond_c) THEN
    channel_fault_c := channel_fault_c + 1;
END_IF;
IF (raw_085_d > 105) AND (NOT cond_d) THEN
    channel_fault_d := channel_fault_d + 1;
END_IF;
IF vote_ok AND train_a_inhibit THEN
    diagnosis_count := diagnosis_count + 1;
END_IF;
IF vote_ok AND train_b_inhibit THEN
    diagnosis_count := diagnosis_count + 1;
END_IF;

cond_a := LimitHigh(raw_086_a, 106);
cond_a := cond_a AND quality_a;
cond_a := cond_a AND (NOT bypass_a);
input_valid_a := InputValid(raw_086_a, 0, 1000);
cond_a := cond_a AND input_valid_a;
IF NOT input_valid_a THEN
    channel_fault_a := channel_fault_a + 1;
END_IF;
cond_b := LimitHigh(raw_086_b, 106);
cond_b := cond_b AND quality_b;
cond_b := cond_b AND (NOT bypass_b);
input_valid_b := InputValid(raw_086_b, 0, 1000);
cond_b := cond_b AND input_valid_b;
IF NOT input_valid_b THEN
    channel_fault_b := channel_fault_b + 1;
END_IF;
cond_c := LimitHigh(raw_086_c, 106);
cond_c := cond_c AND quality_c;
cond_c := cond_c AND (NOT bypass_c);
input_valid_c := InputValid(raw_086_c, 0, 1000);
cond_c := cond_c AND input_valid_c;
IF NOT input_valid_c THEN
    channel_fault_c := channel_fault_c + 1;
END_IF;
cond_d := LimitHigh(raw_086_d, 106);
cond_d := cond_d AND quality_d;
cond_d := cond_d AND (NOT bypass_d);
input_valid_d := InputValid(raw_086_d, 0, 1000);
cond_d := cond_d AND input_valid_d;
IF NOT input_valid_d THEN
    channel_fault_d := channel_fault_d + 1;
END_IF;
vote_ok := TwoOfFour(cond_a, cond_b, cond_c, cond_d);
IF cond_a <> cond_b THEN
    diagnosis_count := diagnosis_count + 1;
END_IF;
IF cond_c <> cond_d THEN
    diagnosis_count := diagnosis_count + 1;
END_IF;
IF NOT vote_ok THEN
    diagnosis_count := diagnosis_count + 1;
END_IF;
latch_a_086 := RS_Next(vote_ok, train_a_reset, latch_a_086);
IF latch_a_086 AND (NOT train_a_inhibit) THEN
    mask_a_10 := mask_a_10 + 64;
    trip_a := 0 < 1;
    scram_a := 0 < 1;
    breaker_a := 0 > 1;
    mfw_a := 0 < 1;
    alarm_a := 0 < 1;
END_IF;
latch_b_086 := RS_Next(vote_ok, train_b_reset, latch_b_086);
IF latch_b_086 AND (NOT train_b_inhibit) THEN
    mask_b_10 := mask_b_10 + 64;
    trip_b := 0 < 1;
    scram_b := 0 < 1;
    breaker_b := 0 > 1;
    mfw_b := 0 < 1;
    alarm_b := 0 < 1;
END_IF;
IF (raw_086_a > 106) AND (NOT cond_a) THEN
    channel_fault_a := channel_fault_a + 1;
END_IF;
IF (raw_086_b > 106) AND (NOT cond_b) THEN
    channel_fault_b := channel_fault_b + 1;
END_IF;
IF (raw_086_c > 106) AND (NOT cond_c) THEN
    channel_fault_c := channel_fault_c + 1;
END_IF;
IF (raw_086_d > 106) AND (NOT cond_d) THEN
    channel_fault_d := channel_fault_d + 1;
END_IF;
IF vote_ok AND train_a_inhibit THEN
    diagnosis_count := diagnosis_count + 1;
END_IF;
IF vote_ok AND train_b_inhibit THEN
    diagnosis_count := diagnosis_count + 1;
END_IF;

cond_a := LimitHigh(raw_087_a, 107);
cond_a := cond_a AND quality_a;
cond_a := cond_a AND (NOT bypass_a);
input_valid_a := InputValid(raw_087_a, 0, 1000);
cond_a := cond_a AND input_valid_a;
IF NOT input_valid_a THEN
    channel_fault_a := channel_fault_a + 1;
END_IF;
cond_b := LimitHigh(raw_087_b, 107);
cond_b := cond_b AND quality_b;
cond_b := cond_b AND (NOT bypass_b);
input_valid_b := InputValid(raw_087_b, 0, 1000);
cond_b := cond_b AND input_valid_b;
IF NOT input_valid_b THEN
    channel_fault_b := channel_fault_b + 1;
END_IF;
cond_c := LimitHigh(raw_087_c, 107);
cond_c := cond_c AND quality_c;
cond_c := cond_c AND (NOT bypass_c);
input_valid_c := InputValid(raw_087_c, 0, 1000);
cond_c := cond_c AND input_valid_c;
IF NOT input_valid_c THEN
    channel_fault_c := channel_fault_c + 1;
END_IF;
cond_d := LimitHigh(raw_087_d, 107);
cond_d := cond_d AND quality_d;
cond_d := cond_d AND (NOT bypass_d);
input_valid_d := InputValid(raw_087_d, 0, 1000);
cond_d := cond_d AND input_valid_d;
IF NOT input_valid_d THEN
    channel_fault_d := channel_fault_d + 1;
END_IF;
vote_ok := TwoOfFour(cond_a, cond_b, cond_c, cond_d);
IF cond_a <> cond_b THEN
    diagnosis_count := diagnosis_count + 1;
END_IF;
IF cond_c <> cond_d THEN
    diagnosis_count := diagnosis_count + 1;
END_IF;
IF NOT vote_ok THEN
    diagnosis_count := diagnosis_count + 1;
END_IF;
latch_a_087 := RS_Next(vote_ok, train_a_reset, latch_a_087);
IF latch_a_087 AND (NOT train_a_inhibit) THEN
    mask_a_10 := mask_a_10 + 128;
    trip_a := 0 < 1;
    scram_a := 0 < 1;
    breaker_a := 0 > 1;
    afw_a := 0 < 1;
    alarm_a := 0 < 1;
END_IF;
latch_b_087 := RS_Next(vote_ok, train_b_reset, latch_b_087);
IF latch_b_087 AND (NOT train_b_inhibit) THEN
    mask_b_10 := mask_b_10 + 128;
    trip_b := 0 < 1;
    scram_b := 0 < 1;
    breaker_b := 0 > 1;
    afw_b := 0 < 1;
    alarm_b := 0 < 1;
END_IF;
IF (raw_087_a > 107) AND (NOT cond_a) THEN
    channel_fault_a := channel_fault_a + 1;
END_IF;
IF (raw_087_b > 107) AND (NOT cond_b) THEN
    channel_fault_b := channel_fault_b + 1;
END_IF;
IF (raw_087_c > 107) AND (NOT cond_c) THEN
    channel_fault_c := channel_fault_c + 1;
END_IF;
IF (raw_087_d > 107) AND (NOT cond_d) THEN
    channel_fault_d := channel_fault_d + 1;
END_IF;
IF vote_ok AND train_a_inhibit THEN
    diagnosis_count := diagnosis_count + 1;
END_IF;
IF vote_ok AND train_b_inhibit THEN
    diagnosis_count := diagnosis_count + 1;
END_IF;

cond_a := LimitHigh(raw_088_a, 108);
cond_a := cond_a AND quality_a;
cond_a := cond_a AND (NOT bypass_a);
input_valid_a := InputValid(raw_088_a, 0, 1000);
cond_a := cond_a AND input_valid_a;
IF NOT input_valid_a THEN
    channel_fault_a := channel_fault_a + 1;
END_IF;
cond_b := LimitHigh(raw_088_b, 108);
cond_b := cond_b AND quality_b;
cond_b := cond_b AND (NOT bypass_b);
input_valid_b := InputValid(raw_088_b, 0, 1000);
cond_b := cond_b AND input_valid_b;
IF NOT input_valid_b THEN
    channel_fault_b := channel_fault_b + 1;
END_IF;
cond_c := LimitHigh(raw_088_c, 108);
cond_c := cond_c AND quality_c;
cond_c := cond_c AND (NOT bypass_c);
input_valid_c := InputValid(raw_088_c, 0, 1000);
cond_c := cond_c AND input_valid_c;
IF NOT input_valid_c THEN
    channel_fault_c := channel_fault_c + 1;
END_IF;
cond_d := LimitHigh(raw_088_d, 108);
cond_d := cond_d AND quality_d;
cond_d := cond_d AND (NOT bypass_d);
input_valid_d := InputValid(raw_088_d, 0, 1000);
cond_d := cond_d AND input_valid_d;
IF NOT input_valid_d THEN
    channel_fault_d := channel_fault_d + 1;
END_IF;
vote_ok := TwoOfFour(cond_a, cond_b, cond_c, cond_d);
IF cond_a <> cond_b THEN
    diagnosis_count := diagnosis_count + 1;
END_IF;
IF cond_c <> cond_d THEN
    diagnosis_count := diagnosis_count + 1;
END_IF;
IF NOT vote_ok THEN
    diagnosis_count := diagnosis_count + 1;
END_IF;
latch_a_088 := RS_Next(vote_ok, train_a_reset, latch_a_088);
IF latch_a_088 AND (NOT train_a_inhibit) THEN
    mask_a_11 := mask_a_11 + 1;
    trip_a := 0 < 1;
    scram_a := 0 < 1;
    breaker_a := 0 > 1;
    si_a := 0 < 1;
    alarm_a := 0 < 1;
END_IF;
latch_b_088 := RS_Next(vote_ok, train_b_reset, latch_b_088);
IF latch_b_088 AND (NOT train_b_inhibit) THEN
    mask_b_11 := mask_b_11 + 1;
    trip_b := 0 < 1;
    scram_b := 0 < 1;
    breaker_b := 0 > 1;
    si_b := 0 < 1;
    alarm_b := 0 < 1;
END_IF;
IF (raw_088_a > 108) AND (NOT cond_a) THEN
    channel_fault_a := channel_fault_a + 1;
END_IF;
IF (raw_088_b > 108) AND (NOT cond_b) THEN
    channel_fault_b := channel_fault_b + 1;
END_IF;
IF (raw_088_c > 108) AND (NOT cond_c) THEN
    channel_fault_c := channel_fault_c + 1;
END_IF;
IF (raw_088_d > 108) AND (NOT cond_d) THEN
    channel_fault_d := channel_fault_d + 1;
END_IF;
IF vote_ok AND train_a_inhibit THEN
    diagnosis_count := diagnosis_count + 1;
END_IF;
IF vote_ok AND train_b_inhibit THEN
    diagnosis_count := diagnosis_count + 1;
END_IF;

cond_a := LimitHigh(raw_089_a, 109);
cond_a := cond_a AND quality_a;
cond_a := cond_a AND (NOT bypass_a);
input_valid_a := InputValid(raw_089_a, 0, 1000);
cond_a := cond_a AND input_valid_a;
IF NOT input_valid_a THEN
    channel_fault_a := channel_fault_a + 1;
END_IF;
cond_b := LimitHigh(raw_089_b, 109);
cond_b := cond_b AND quality_b;
cond_b := cond_b AND (NOT bypass_b);
input_valid_b := InputValid(raw_089_b, 0, 1000);
cond_b := cond_b AND input_valid_b;
IF NOT input_valid_b THEN
    channel_fault_b := channel_fault_b + 1;
END_IF;
cond_c := LimitHigh(raw_089_c, 109);
cond_c := cond_c AND quality_c;
cond_c := cond_c AND (NOT bypass_c);
input_valid_c := InputValid(raw_089_c, 0, 1000);
cond_c := cond_c AND input_valid_c;
IF NOT input_valid_c THEN
    channel_fault_c := channel_fault_c + 1;
END_IF;
cond_d := LimitHigh(raw_089_d, 109);
cond_d := cond_d AND quality_d;
cond_d := cond_d AND (NOT bypass_d);
input_valid_d := InputValid(raw_089_d, 0, 1000);
cond_d := cond_d AND input_valid_d;
IF NOT input_valid_d THEN
    channel_fault_d := channel_fault_d + 1;
END_IF;
vote_ok := TwoOfFour(cond_a, cond_b, cond_c, cond_d);
IF cond_a <> cond_b THEN
    diagnosis_count := diagnosis_count + 1;
END_IF;
IF cond_c <> cond_d THEN
    diagnosis_count := diagnosis_count + 1;
END_IF;
IF NOT vote_ok THEN
    diagnosis_count := diagnosis_count + 1;
END_IF;
latch_a_089 := RS_Next(vote_ok, train_a_reset, latch_a_089);
IF latch_a_089 AND (NOT train_a_inhibit) THEN
    mask_a_11 := mask_a_11 + 2;
    trip_a := 0 < 1;
    scram_a := 0 < 1;
    breaker_a := 0 > 1;
    ci_a := 0 < 1;
    alarm_a := 0 < 1;
END_IF;
latch_b_089 := RS_Next(vote_ok, train_b_reset, latch_b_089);
IF latch_b_089 AND (NOT train_b_inhibit) THEN
    mask_b_11 := mask_b_11 + 2;
    trip_b := 0 < 1;
    scram_b := 0 < 1;
    breaker_b := 0 > 1;
    ci_b := 0 < 1;
    alarm_b := 0 < 1;
END_IF;
IF (raw_089_a > 109) AND (NOT cond_a) THEN
    channel_fault_a := channel_fault_a + 1;
END_IF;
IF (raw_089_b > 109) AND (NOT cond_b) THEN
    channel_fault_b := channel_fault_b + 1;
END_IF;
IF (raw_089_c > 109) AND (NOT cond_c) THEN
    channel_fault_c := channel_fault_c + 1;
END_IF;
IF (raw_089_d > 109) AND (NOT cond_d) THEN
    channel_fault_d := channel_fault_d + 1;
END_IF;
IF vote_ok AND train_a_inhibit THEN
    diagnosis_count := diagnosis_count + 1;
END_IF;
IF vote_ok AND train_b_inhibit THEN
    diagnosis_count := diagnosis_count + 1;
END_IF;

cond_a := LimitHigh(raw_090_a, 110);
cond_a := cond_a AND quality_a;
cond_a := cond_a AND (NOT bypass_a);
input_valid_a := InputValid(raw_090_a, 0, 1000);
cond_a := cond_a AND input_valid_a;
IF NOT input_valid_a THEN
    channel_fault_a := channel_fault_a + 1;
END_IF;
cond_b := LimitHigh(raw_090_b, 110);
cond_b := cond_b AND quality_b;
cond_b := cond_b AND (NOT bypass_b);
input_valid_b := InputValid(raw_090_b, 0, 1000);
cond_b := cond_b AND input_valid_b;
IF NOT input_valid_b THEN
    channel_fault_b := channel_fault_b + 1;
END_IF;
cond_c := LimitHigh(raw_090_c, 110);
cond_c := cond_c AND quality_c;
cond_c := cond_c AND (NOT bypass_c);
input_valid_c := InputValid(raw_090_c, 0, 1000);
cond_c := cond_c AND input_valid_c;
IF NOT input_valid_c THEN
    channel_fault_c := channel_fault_c + 1;
END_IF;
cond_d := LimitHigh(raw_090_d, 110);
cond_d := cond_d AND quality_d;
cond_d := cond_d AND (NOT bypass_d);
input_valid_d := InputValid(raw_090_d, 0, 1000);
cond_d := cond_d AND input_valid_d;
IF NOT input_valid_d THEN
    channel_fault_d := channel_fault_d + 1;
END_IF;
vote_ok := TwoOfFour(cond_a, cond_b, cond_c, cond_d);
IF cond_a <> cond_b THEN
    diagnosis_count := diagnosis_count + 1;
END_IF;
IF cond_c <> cond_d THEN
    diagnosis_count := diagnosis_count + 1;
END_IF;
IF NOT vote_ok THEN
    diagnosis_count := diagnosis_count + 1;
END_IF;
latch_a_090 := RS_Next(vote_ok, train_a_reset, latch_a_090);
IF latch_a_090 AND (NOT train_a_inhibit) THEN
    mask_a_11 := mask_a_11 + 4;
    trip_a := 0 < 1;
    scram_a := 0 < 1;
    breaker_a := 0 > 1;
    mfw_a := 0 < 1;
    alarm_a := 0 < 1;
END_IF;
latch_b_090 := RS_Next(vote_ok, train_b_reset, latch_b_090);
IF latch_b_090 AND (NOT train_b_inhibit) THEN
    mask_b_11 := mask_b_11 + 4;
    trip_b := 0 < 1;
    scram_b := 0 < 1;
    breaker_b := 0 > 1;
    mfw_b := 0 < 1;
    alarm_b := 0 < 1;
END_IF;
IF (raw_090_a > 110) AND (NOT cond_a) THEN
    channel_fault_a := channel_fault_a + 1;
END_IF;
IF (raw_090_b > 110) AND (NOT cond_b) THEN
    channel_fault_b := channel_fault_b + 1;
END_IF;
IF (raw_090_c > 110) AND (NOT cond_c) THEN
    channel_fault_c := channel_fault_c + 1;
END_IF;
IF (raw_090_d > 110) AND (NOT cond_d) THEN
    channel_fault_d := channel_fault_d + 1;
END_IF;
IF vote_ok AND train_a_inhibit THEN
    diagnosis_count := diagnosis_count + 1;
END_IF;
IF vote_ok AND train_b_inhibit THEN
    diagnosis_count := diagnosis_count + 1;
END_IF;

cond_a := LimitHigh(raw_091_a, 111);
cond_a := cond_a AND quality_a;
cond_a := cond_a AND (NOT bypass_a);
input_valid_a := InputValid(raw_091_a, 0, 1000);
cond_a := cond_a AND input_valid_a;
IF NOT input_valid_a THEN
    channel_fault_a := channel_fault_a + 1;
END_IF;
cond_b := LimitHigh(raw_091_b, 111);
cond_b := cond_b AND quality_b;
cond_b := cond_b AND (NOT bypass_b);
input_valid_b := InputValid(raw_091_b, 0, 1000);
cond_b := cond_b AND input_valid_b;
IF NOT input_valid_b THEN
    channel_fault_b := channel_fault_b + 1;
END_IF;
cond_c := LimitHigh(raw_091_c, 111);
cond_c := cond_c AND quality_c;
cond_c := cond_c AND (NOT bypass_c);
input_valid_c := InputValid(raw_091_c, 0, 1000);
cond_c := cond_c AND input_valid_c;
IF NOT input_valid_c THEN
    channel_fault_c := channel_fault_c + 1;
END_IF;
cond_d := LimitHigh(raw_091_d, 111);
cond_d := cond_d AND quality_d;
cond_d := cond_d AND (NOT bypass_d);
input_valid_d := InputValid(raw_091_d, 0, 1000);
cond_d := cond_d AND input_valid_d;
IF NOT input_valid_d THEN
    channel_fault_d := channel_fault_d + 1;
END_IF;
vote_ok := TwoOfFour(cond_a, cond_b, cond_c, cond_d);
IF cond_a <> cond_b THEN
    diagnosis_count := diagnosis_count + 1;
END_IF;
IF cond_c <> cond_d THEN
    diagnosis_count := diagnosis_count + 1;
END_IF;
IF NOT vote_ok THEN
    diagnosis_count := diagnosis_count + 1;
END_IF;
latch_a_091 := RS_Next(vote_ok, train_a_reset, latch_a_091);
IF latch_a_091 AND (NOT train_a_inhibit) THEN
    mask_a_11 := mask_a_11 + 8;
    trip_a := 0 < 1;
    scram_a := 0 < 1;
    breaker_a := 0 > 1;
    afw_a := 0 < 1;
    alarm_a := 0 < 1;
END_IF;
latch_b_091 := RS_Next(vote_ok, train_b_reset, latch_b_091);
IF latch_b_091 AND (NOT train_b_inhibit) THEN
    mask_b_11 := mask_b_11 + 8;
    trip_b := 0 < 1;
    scram_b := 0 < 1;
    breaker_b := 0 > 1;
    afw_b := 0 < 1;
    alarm_b := 0 < 1;
END_IF;
IF (raw_091_a > 111) AND (NOT cond_a) THEN
    channel_fault_a := channel_fault_a + 1;
END_IF;
IF (raw_091_b > 111) AND (NOT cond_b) THEN
    channel_fault_b := channel_fault_b + 1;
END_IF;
IF (raw_091_c > 111) AND (NOT cond_c) THEN
    channel_fault_c := channel_fault_c + 1;
END_IF;
IF (raw_091_d > 111) AND (NOT cond_d) THEN
    channel_fault_d := channel_fault_d + 1;
END_IF;
IF vote_ok AND train_a_inhibit THEN
    diagnosis_count := diagnosis_count + 1;
END_IF;
IF vote_ok AND train_b_inhibit THEN
    diagnosis_count := diagnosis_count + 1;
END_IF;

cond_a := LimitHigh(raw_092_a, 112);
cond_a := cond_a AND quality_a;
cond_a := cond_a AND (NOT bypass_a);
input_valid_a := InputValid(raw_092_a, 0, 1000);
cond_a := cond_a AND input_valid_a;
IF NOT input_valid_a THEN
    channel_fault_a := channel_fault_a + 1;
END_IF;
cond_b := LimitHigh(raw_092_b, 112);
cond_b := cond_b AND quality_b;
cond_b := cond_b AND (NOT bypass_b);
input_valid_b := InputValid(raw_092_b, 0, 1000);
cond_b := cond_b AND input_valid_b;
IF NOT input_valid_b THEN
    channel_fault_b := channel_fault_b + 1;
END_IF;
cond_c := LimitHigh(raw_092_c, 112);
cond_c := cond_c AND quality_c;
cond_c := cond_c AND (NOT bypass_c);
input_valid_c := InputValid(raw_092_c, 0, 1000);
cond_c := cond_c AND input_valid_c;
IF NOT input_valid_c THEN
    channel_fault_c := channel_fault_c + 1;
END_IF;
cond_d := LimitHigh(raw_092_d, 112);
cond_d := cond_d AND quality_d;
cond_d := cond_d AND (NOT bypass_d);
input_valid_d := InputValid(raw_092_d, 0, 1000);
cond_d := cond_d AND input_valid_d;
IF NOT input_valid_d THEN
    channel_fault_d := channel_fault_d + 1;
END_IF;
vote_ok := TwoOfFour(cond_a, cond_b, cond_c, cond_d);
IF cond_a <> cond_b THEN
    diagnosis_count := diagnosis_count + 1;
END_IF;
IF cond_c <> cond_d THEN
    diagnosis_count := diagnosis_count + 1;
END_IF;
IF NOT vote_ok THEN
    diagnosis_count := diagnosis_count + 1;
END_IF;
latch_a_092 := RS_Next(vote_ok, train_a_reset, latch_a_092);
IF latch_a_092 AND (NOT train_a_inhibit) THEN
    mask_a_11 := mask_a_11 + 16;
    trip_a := 0 < 1;
    scram_a := 0 < 1;
    breaker_a := 0 > 1;
    si_a := 0 < 1;
    alarm_a := 0 < 1;
END_IF;
latch_b_092 := RS_Next(vote_ok, train_b_reset, latch_b_092);
IF latch_b_092 AND (NOT train_b_inhibit) THEN
    mask_b_11 := mask_b_11 + 16;
    trip_b := 0 < 1;
    scram_b := 0 < 1;
    breaker_b := 0 > 1;
    si_b := 0 < 1;
    alarm_b := 0 < 1;
END_IF;
IF (raw_092_a > 112) AND (NOT cond_a) THEN
    channel_fault_a := channel_fault_a + 1;
END_IF;
IF (raw_092_b > 112) AND (NOT cond_b) THEN
    channel_fault_b := channel_fault_b + 1;
END_IF;
IF (raw_092_c > 112) AND (NOT cond_c) THEN
    channel_fault_c := channel_fault_c + 1;
END_IF;
IF (raw_092_d > 112) AND (NOT cond_d) THEN
    channel_fault_d := channel_fault_d + 1;
END_IF;
IF vote_ok AND train_a_inhibit THEN
    diagnosis_count := diagnosis_count + 1;
END_IF;
IF vote_ok AND train_b_inhibit THEN
    diagnosis_count := diagnosis_count + 1;
END_IF;

cond_a := LimitHigh(raw_093_a, 113);
cond_a := cond_a AND quality_a;
cond_a := cond_a AND (NOT bypass_a);
input_valid_a := InputValid(raw_093_a, 0, 1000);
cond_a := cond_a AND input_valid_a;
IF NOT input_valid_a THEN
    channel_fault_a := channel_fault_a + 1;
END_IF;
cond_b := LimitHigh(raw_093_b, 113);
cond_b := cond_b AND quality_b;
cond_b := cond_b AND (NOT bypass_b);
input_valid_b := InputValid(raw_093_b, 0, 1000);
cond_b := cond_b AND input_valid_b;
IF NOT input_valid_b THEN
    channel_fault_b := channel_fault_b + 1;
END_IF;
cond_c := LimitHigh(raw_093_c, 113);
cond_c := cond_c AND quality_c;
cond_c := cond_c AND (NOT bypass_c);
input_valid_c := InputValid(raw_093_c, 0, 1000);
cond_c := cond_c AND input_valid_c;
IF NOT input_valid_c THEN
    channel_fault_c := channel_fault_c + 1;
END_IF;
cond_d := LimitHigh(raw_093_d, 113);
cond_d := cond_d AND quality_d;
cond_d := cond_d AND (NOT bypass_d);
input_valid_d := InputValid(raw_093_d, 0, 1000);
cond_d := cond_d AND input_valid_d;
IF NOT input_valid_d THEN
    channel_fault_d := channel_fault_d + 1;
END_IF;
vote_ok := TwoOfFour(cond_a, cond_b, cond_c, cond_d);
IF cond_a <> cond_b THEN
    diagnosis_count := diagnosis_count + 1;
END_IF;
IF cond_c <> cond_d THEN
    diagnosis_count := diagnosis_count + 1;
END_IF;
IF NOT vote_ok THEN
    diagnosis_count := diagnosis_count + 1;
END_IF;
latch_a_093 := RS_Next(vote_ok, train_a_reset, latch_a_093);
IF latch_a_093 AND (NOT train_a_inhibit) THEN
    mask_a_11 := mask_a_11 + 32;
    trip_a := 0 < 1;
    scram_a := 0 < 1;
    breaker_a := 0 > 1;
    ci_a := 0 < 1;
    alarm_a := 0 < 1;
END_IF;
latch_b_093 := RS_Next(vote_ok, train_b_reset, latch_b_093);
IF latch_b_093 AND (NOT train_b_inhibit) THEN
    mask_b_11 := mask_b_11 + 32;
    trip_b := 0 < 1;
    scram_b := 0 < 1;
    breaker_b := 0 > 1;
    ci_b := 0 < 1;
    alarm_b := 0 < 1;
END_IF;
IF (raw_093_a > 113) AND (NOT cond_a) THEN
    channel_fault_a := channel_fault_a + 1;
END_IF;
IF (raw_093_b > 113) AND (NOT cond_b) THEN
    channel_fault_b := channel_fault_b + 1;
END_IF;
IF (raw_093_c > 113) AND (NOT cond_c) THEN
    channel_fault_c := channel_fault_c + 1;
END_IF;
IF (raw_093_d > 113) AND (NOT cond_d) THEN
    channel_fault_d := channel_fault_d + 1;
END_IF;
IF vote_ok AND train_a_inhibit THEN
    diagnosis_count := diagnosis_count + 1;
END_IF;
IF vote_ok AND train_b_inhibit THEN
    diagnosis_count := diagnosis_count + 1;
END_IF;

cond_a := LimitHigh(raw_094_a, 114);
cond_a := cond_a AND quality_a;
cond_a := cond_a AND (NOT bypass_a);
input_valid_a := InputValid(raw_094_a, 0, 1000);
cond_a := cond_a AND input_valid_a;
IF NOT input_valid_a THEN
    channel_fault_a := channel_fault_a + 1;
END_IF;
cond_b := LimitHigh(raw_094_b, 114);
cond_b := cond_b AND quality_b;
cond_b := cond_b AND (NOT bypass_b);
input_valid_b := InputValid(raw_094_b, 0, 1000);
cond_b := cond_b AND input_valid_b;
IF NOT input_valid_b THEN
    channel_fault_b := channel_fault_b + 1;
END_IF;
cond_c := LimitHigh(raw_094_c, 114);
cond_c := cond_c AND quality_c;
cond_c := cond_c AND (NOT bypass_c);
input_valid_c := InputValid(raw_094_c, 0, 1000);
cond_c := cond_c AND input_valid_c;
IF NOT input_valid_c THEN
    channel_fault_c := channel_fault_c + 1;
END_IF;
cond_d := LimitHigh(raw_094_d, 114);
cond_d := cond_d AND quality_d;
cond_d := cond_d AND (NOT bypass_d);
input_valid_d := InputValid(raw_094_d, 0, 1000);
cond_d := cond_d AND input_valid_d;
IF NOT input_valid_d THEN
    channel_fault_d := channel_fault_d + 1;
END_IF;
vote_ok := TwoOfFour(cond_a, cond_b, cond_c, cond_d);
IF cond_a <> cond_b THEN
    diagnosis_count := diagnosis_count + 1;
END_IF;
IF cond_c <> cond_d THEN
    diagnosis_count := diagnosis_count + 1;
END_IF;
IF NOT vote_ok THEN
    diagnosis_count := diagnosis_count + 1;
END_IF;
latch_a_094 := RS_Next(vote_ok, train_a_reset, latch_a_094);
IF latch_a_094 AND (NOT train_a_inhibit) THEN
    mask_a_11 := mask_a_11 + 64;
    trip_a := 0 < 1;
    scram_a := 0 < 1;
    breaker_a := 0 > 1;
    mfw_a := 0 < 1;
    alarm_a := 0 < 1;
END_IF;
latch_b_094 := RS_Next(vote_ok, train_b_reset, latch_b_094);
IF latch_b_094 AND (NOT train_b_inhibit) THEN
    mask_b_11 := mask_b_11 + 64;
    trip_b := 0 < 1;
    scram_b := 0 < 1;
    breaker_b := 0 > 1;
    mfw_b := 0 < 1;
    alarm_b := 0 < 1;
END_IF;
IF (raw_094_a > 114) AND (NOT cond_a) THEN
    channel_fault_a := channel_fault_a + 1;
END_IF;
IF (raw_094_b > 114) AND (NOT cond_b) THEN
    channel_fault_b := channel_fault_b + 1;
END_IF;
IF (raw_094_c > 114) AND (NOT cond_c) THEN
    channel_fault_c := channel_fault_c + 1;
END_IF;
IF (raw_094_d > 114) AND (NOT cond_d) THEN
    channel_fault_d := channel_fault_d + 1;
END_IF;
IF vote_ok AND train_a_inhibit THEN
    diagnosis_count := diagnosis_count + 1;
END_IF;
IF vote_ok AND train_b_inhibit THEN
    diagnosis_count := diagnosis_count + 1;
END_IF;

cond_a := LimitHigh(raw_095_a, 115);
cond_a := cond_a AND quality_a;
cond_a := cond_a AND (NOT bypass_a);
input_valid_a := InputValid(raw_095_a, 0, 1000);
cond_a := cond_a AND input_valid_a;
IF NOT input_valid_a THEN
    channel_fault_a := channel_fault_a + 1;
END_IF;
cond_b := LimitHigh(raw_095_b, 115);
cond_b := cond_b AND quality_b;
cond_b := cond_b AND (NOT bypass_b);
input_valid_b := InputValid(raw_095_b, 0, 1000);
cond_b := cond_b AND input_valid_b;
IF NOT input_valid_b THEN
    channel_fault_b := channel_fault_b + 1;
END_IF;
cond_c := LimitHigh(raw_095_c, 115);
cond_c := cond_c AND quality_c;
cond_c := cond_c AND (NOT bypass_c);
input_valid_c := InputValid(raw_095_c, 0, 1000);
cond_c := cond_c AND input_valid_c;
IF NOT input_valid_c THEN
    channel_fault_c := channel_fault_c + 1;
END_IF;
cond_d := LimitHigh(raw_095_d, 115);
cond_d := cond_d AND quality_d;
cond_d := cond_d AND (NOT bypass_d);
input_valid_d := InputValid(raw_095_d, 0, 1000);
cond_d := cond_d AND input_valid_d;
IF NOT input_valid_d THEN
    channel_fault_d := channel_fault_d + 1;
END_IF;
vote_ok := TwoOfFour(cond_a, cond_b, cond_c, cond_d);
IF cond_a <> cond_b THEN
    diagnosis_count := diagnosis_count + 1;
END_IF;
IF cond_c <> cond_d THEN
    diagnosis_count := diagnosis_count + 1;
END_IF;
IF NOT vote_ok THEN
    diagnosis_count := diagnosis_count + 1;
END_IF;
latch_a_095 := RS_Next(vote_ok, train_a_reset, latch_a_095);
IF latch_a_095 AND (NOT train_a_inhibit) THEN
    mask_a_11 := mask_a_11 + 128;
    trip_a := 0 < 1;
    scram_a := 0 < 1;
    breaker_a := 0 > 1;
    afw_a := 0 < 1;
    alarm_a := 0 < 1;
END_IF;
latch_b_095 := RS_Next(vote_ok, train_b_reset, latch_b_095);
IF latch_b_095 AND (NOT train_b_inhibit) THEN
    mask_b_11 := mask_b_11 + 128;
    trip_b := 0 < 1;
    scram_b := 0 < 1;
    breaker_b := 0 > 1;
    afw_b := 0 < 1;
    alarm_b := 0 < 1;
END_IF;
IF (raw_095_a > 115) AND (NOT cond_a) THEN
    channel_fault_a := channel_fault_a + 1;
END_IF;
IF (raw_095_b > 115) AND (NOT cond_b) THEN
    channel_fault_b := channel_fault_b + 1;
END_IF;
IF (raw_095_c > 115) AND (NOT cond_c) THEN
    channel_fault_c := channel_fault_c + 1;
END_IF;
IF (raw_095_d > 115) AND (NOT cond_d) THEN
    channel_fault_d := channel_fault_d + 1;
END_IF;
IF vote_ok AND train_a_inhibit THEN
    diagnosis_count := diagnosis_count + 1;
END_IF;
IF vote_ok AND train_b_inhibit THEN
    diagnosis_count := diagnosis_count + 1;
END_IF;

cond_a := LimitHigh(raw_096_a, 116);
cond_a := cond_a AND quality_a;
cond_a := cond_a AND (NOT bypass_a);
input_valid_a := InputValid(raw_096_a, 0, 1000);
cond_a := cond_a AND input_valid_a;
IF NOT input_valid_a THEN
    channel_fault_a := channel_fault_a + 1;
END_IF;
cond_b := LimitHigh(raw_096_b, 116);
cond_b := cond_b AND quality_b;
cond_b := cond_b AND (NOT bypass_b);
input_valid_b := InputValid(raw_096_b, 0, 1000);
cond_b := cond_b AND input_valid_b;
IF NOT input_valid_b THEN
    channel_fault_b := channel_fault_b + 1;
END_IF;
cond_c := LimitHigh(raw_096_c, 116);
cond_c := cond_c AND quality_c;
cond_c := cond_c AND (NOT bypass_c);
input_valid_c := InputValid(raw_096_c, 0, 1000);
cond_c := cond_c AND input_valid_c;
IF NOT input_valid_c THEN
    channel_fault_c := channel_fault_c + 1;
END_IF;
cond_d := LimitHigh(raw_096_d, 116);
cond_d := cond_d AND quality_d;
cond_d := cond_d AND (NOT bypass_d);
input_valid_d := InputValid(raw_096_d, 0, 1000);
cond_d := cond_d AND input_valid_d;
IF NOT input_valid_d THEN
    channel_fault_d := channel_fault_d + 1;
END_IF;
vote_ok := TwoOfFour(cond_a, cond_b, cond_c, cond_d);
IF cond_a <> cond_b THEN
    diagnosis_count := diagnosis_count + 1;
END_IF;
IF cond_c <> cond_d THEN
    diagnosis_count := diagnosis_count + 1;
END_IF;
IF NOT vote_ok THEN
    diagnosis_count := diagnosis_count + 1;
END_IF;
latch_a_096 := RS_Next(vote_ok, train_a_reset, latch_a_096);
IF latch_a_096 AND (NOT train_a_inhibit) THEN
    mask_a_12 := mask_a_12 + 1;
    trip_a := 0 < 1;
    scram_a := 0 < 1;
    breaker_a := 0 > 1;
    si_a := 0 < 1;
    alarm_a := 0 < 1;
END_IF;
latch_b_096 := RS_Next(vote_ok, train_b_reset, latch_b_096);
IF latch_b_096 AND (NOT train_b_inhibit) THEN
    mask_b_12 := mask_b_12 + 1;
    trip_b := 0 < 1;
    scram_b := 0 < 1;
    breaker_b := 0 > 1;
    si_b := 0 < 1;
    alarm_b := 0 < 1;
END_IF;
IF (raw_096_a > 116) AND (NOT cond_a) THEN
    channel_fault_a := channel_fault_a + 1;
END_IF;
IF (raw_096_b > 116) AND (NOT cond_b) THEN
    channel_fault_b := channel_fault_b + 1;
END_IF;
IF (raw_096_c > 116) AND (NOT cond_c) THEN
    channel_fault_c := channel_fault_c + 1;
END_IF;
IF (raw_096_d > 116) AND (NOT cond_d) THEN
    channel_fault_d := channel_fault_d + 1;
END_IF;
IF vote_ok AND train_a_inhibit THEN
    diagnosis_count := diagnosis_count + 1;
END_IF;
IF vote_ok AND train_b_inhibit THEN
    diagnosis_count := diagnosis_count + 1;
END_IF;

cond_a := LimitHigh(raw_097_a, 117);
cond_a := cond_a AND quality_a;
cond_a := cond_a AND (NOT bypass_a);
input_valid_a := InputValid(raw_097_a, 0, 1000);
cond_a := cond_a AND input_valid_a;
IF NOT input_valid_a THEN
    channel_fault_a := channel_fault_a + 1;
END_IF;
cond_b := LimitHigh(raw_097_b, 117);
cond_b := cond_b AND quality_b;
cond_b := cond_b AND (NOT bypass_b);
input_valid_b := InputValid(raw_097_b, 0, 1000);
cond_b := cond_b AND input_valid_b;
IF NOT input_valid_b THEN
    channel_fault_b := channel_fault_b + 1;
END_IF;
cond_c := LimitHigh(raw_097_c, 117);
cond_c := cond_c AND quality_c;
cond_c := cond_c AND (NOT bypass_c);
input_valid_c := InputValid(raw_097_c, 0, 1000);
cond_c := cond_c AND input_valid_c;
IF NOT input_valid_c THEN
    channel_fault_c := channel_fault_c + 1;
END_IF;
cond_d := LimitHigh(raw_097_d, 117);
cond_d := cond_d AND quality_d;
cond_d := cond_d AND (NOT bypass_d);
input_valid_d := InputValid(raw_097_d, 0, 1000);
cond_d := cond_d AND input_valid_d;
IF NOT input_valid_d THEN
    channel_fault_d := channel_fault_d + 1;
END_IF;
vote_ok := TwoOfFour(cond_a, cond_b, cond_c, cond_d);
IF cond_a <> cond_b THEN
    diagnosis_count := diagnosis_count + 1;
END_IF;
IF cond_c <> cond_d THEN
    diagnosis_count := diagnosis_count + 1;
END_IF;
IF NOT vote_ok THEN
    diagnosis_count := diagnosis_count + 1;
END_IF;
latch_a_097 := RS_Next(vote_ok, train_a_reset, latch_a_097);
IF latch_a_097 AND (NOT train_a_inhibit) THEN
    mask_a_12 := mask_a_12 + 2;
    trip_a := 0 < 1;
    scram_a := 0 < 1;
    breaker_a := 0 > 1;
    ci_a := 0 < 1;
    alarm_a := 0 < 1;
END_IF;
latch_b_097 := RS_Next(vote_ok, train_b_reset, latch_b_097);
IF latch_b_097 AND (NOT train_b_inhibit) THEN
    mask_b_12 := mask_b_12 + 2;
    trip_b := 0 < 1;
    scram_b := 0 < 1;
    breaker_b := 0 > 1;
    ci_b := 0 < 1;
    alarm_b := 0 < 1;
END_IF;
IF (raw_097_a > 117) AND (NOT cond_a) THEN
    channel_fault_a := channel_fault_a + 1;
END_IF;
IF (raw_097_b > 117) AND (NOT cond_b) THEN
    channel_fault_b := channel_fault_b + 1;
END_IF;
IF (raw_097_c > 117) AND (NOT cond_c) THEN
    channel_fault_c := channel_fault_c + 1;
END_IF;
IF (raw_097_d > 117) AND (NOT cond_d) THEN
    channel_fault_d := channel_fault_d + 1;
END_IF;
IF vote_ok AND train_a_inhibit THEN
    diagnosis_count := diagnosis_count + 1;
END_IF;
IF vote_ok AND train_b_inhibit THEN
    diagnosis_count := diagnosis_count + 1;
END_IF;

cond_a := LimitHigh(raw_098_a, 118);
cond_a := cond_a AND quality_a;
cond_a := cond_a AND (NOT bypass_a);
input_valid_a := InputValid(raw_098_a, 0, 1000);
cond_a := cond_a AND input_valid_a;
IF NOT input_valid_a THEN
    channel_fault_a := channel_fault_a + 1;
END_IF;
cond_b := LimitHigh(raw_098_b, 118);
cond_b := cond_b AND quality_b;
cond_b := cond_b AND (NOT bypass_b);
input_valid_b := InputValid(raw_098_b, 0, 1000);
cond_b := cond_b AND input_valid_b;
IF NOT input_valid_b THEN
    channel_fault_b := channel_fault_b + 1;
END_IF;
cond_c := LimitHigh(raw_098_c, 118);
cond_c := cond_c AND quality_c;
cond_c := cond_c AND (NOT bypass_c);
input_valid_c := InputValid(raw_098_c, 0, 1000);
cond_c := cond_c AND input_valid_c;
IF NOT input_valid_c THEN
    channel_fault_c := channel_fault_c + 1;
END_IF;
cond_d := LimitHigh(raw_098_d, 118);
cond_d := cond_d AND quality_d;
cond_d := cond_d AND (NOT bypass_d);
input_valid_d := InputValid(raw_098_d, 0, 1000);
cond_d := cond_d AND input_valid_d;
IF NOT input_valid_d THEN
    channel_fault_d := channel_fault_d + 1;
END_IF;
vote_ok := TwoOfFour(cond_a, cond_b, cond_c, cond_d);
IF cond_a <> cond_b THEN
    diagnosis_count := diagnosis_count + 1;
END_IF;
IF cond_c <> cond_d THEN
    diagnosis_count := diagnosis_count + 1;
END_IF;
IF NOT vote_ok THEN
    diagnosis_count := diagnosis_count + 1;
END_IF;
latch_a_098 := RS_Next(vote_ok, train_a_reset, latch_a_098);
IF latch_a_098 AND (NOT train_a_inhibit) THEN
    mask_a_12 := mask_a_12 + 4;
    trip_a := 0 < 1;
    scram_a := 0 < 1;
    breaker_a := 0 > 1;
    mfw_a := 0 < 1;
    alarm_a := 0 < 1;
END_IF;
latch_b_098 := RS_Next(vote_ok, train_b_reset, latch_b_098);
IF latch_b_098 AND (NOT train_b_inhibit) THEN
    mask_b_12 := mask_b_12 + 4;
    trip_b := 0 < 1;
    scram_b := 0 < 1;
    breaker_b := 0 > 1;
    mfw_b := 0 < 1;
    alarm_b := 0 < 1;
END_IF;
IF (raw_098_a > 118) AND (NOT cond_a) THEN
    channel_fault_a := channel_fault_a + 1;
END_IF;
IF (raw_098_b > 118) AND (NOT cond_b) THEN
    channel_fault_b := channel_fault_b + 1;
END_IF;
IF (raw_098_c > 118) AND (NOT cond_c) THEN
    channel_fault_c := channel_fault_c + 1;
END_IF;
IF (raw_098_d > 118) AND (NOT cond_d) THEN
    channel_fault_d := channel_fault_d + 1;
END_IF;
IF vote_ok AND train_a_inhibit THEN
    diagnosis_count := diagnosis_count + 1;
END_IF;
IF vote_ok AND train_b_inhibit THEN
    diagnosis_count := diagnosis_count + 1;
END_IF;

cond_a := LimitHigh(raw_099_a, 119);
cond_a := cond_a AND quality_a;
cond_a := cond_a AND (NOT bypass_a);
input_valid_a := InputValid(raw_099_a, 0, 1000);
cond_a := cond_a AND input_valid_a;
IF NOT input_valid_a THEN
    channel_fault_a := channel_fault_a + 1;
END_IF;
cond_b := LimitHigh(raw_099_b, 119);
cond_b := cond_b AND quality_b;
cond_b := cond_b AND (NOT bypass_b);
input_valid_b := InputValid(raw_099_b, 0, 1000);
cond_b := cond_b AND input_valid_b;
IF NOT input_valid_b THEN
    channel_fault_b := channel_fault_b + 1;
END_IF;
cond_c := LimitHigh(raw_099_c, 119);
cond_c := cond_c AND quality_c;
cond_c := cond_c AND (NOT bypass_c);
input_valid_c := InputValid(raw_099_c, 0, 1000);
cond_c := cond_c AND input_valid_c;
IF NOT input_valid_c THEN
    channel_fault_c := channel_fault_c + 1;
END_IF;
cond_d := LimitHigh(raw_099_d, 119);
cond_d := cond_d AND quality_d;
cond_d := cond_d AND (NOT bypass_d);
input_valid_d := InputValid(raw_099_d, 0, 1000);
cond_d := cond_d AND input_valid_d;
IF NOT input_valid_d THEN
    channel_fault_d := channel_fault_d + 1;
END_IF;
vote_ok := TwoOfFour(cond_a, cond_b, cond_c, cond_d);
IF cond_a <> cond_b THEN
    diagnosis_count := diagnosis_count + 1;
END_IF;
IF cond_c <> cond_d THEN
    diagnosis_count := diagnosis_count + 1;
END_IF;
IF NOT vote_ok THEN
    diagnosis_count := diagnosis_count + 1;
END_IF;
latch_a_099 := RS_Next(vote_ok, train_a_reset, latch_a_099);
IF latch_a_099 AND (NOT train_a_inhibit) THEN
    mask_a_12 := mask_a_12 + 8;
    trip_a := 0 < 1;
    scram_a := 0 < 1;
    breaker_a := 0 > 1;
    afw_a := 0 < 1;
    alarm_a := 0 < 1;
END_IF;
latch_b_099 := RS_Next(vote_ok, train_b_reset, latch_b_099);
IF latch_b_099 AND (NOT train_b_inhibit) THEN
    mask_b_12 := mask_b_12 + 8;
    trip_b := 0 < 1;
    scram_b := 0 < 1;
    breaker_b := 0 > 1;
    afw_b := 0 < 1;
    alarm_b := 0 < 1;
END_IF;
IF (raw_099_a > 119) AND (NOT cond_a) THEN
    channel_fault_a := channel_fault_a + 1;
END_IF;
IF (raw_099_b > 119) AND (NOT cond_b) THEN
    channel_fault_b := channel_fault_b + 1;
END_IF;
IF (raw_099_c > 119) AND (NOT cond_c) THEN
    channel_fault_c := channel_fault_c + 1;
END_IF;
IF (raw_099_d > 119) AND (NOT cond_d) THEN
    channel_fault_d := channel_fault_d + 1;
END_IF;
IF vote_ok AND train_a_inhibit THEN
    diagnosis_count := diagnosis_count + 1;
END_IF;
IF vote_ok AND train_b_inhibit THEN
    diagnosis_count := diagnosis_count + 1;
END_IF;

cond_a := LimitHigh(raw_100_a, 120);
cond_a := cond_a AND quality_a;
cond_a := cond_a AND (NOT bypass_a);
input_valid_a := InputValid(raw_100_a, 0, 1000);
cond_a := cond_a AND input_valid_a;
IF NOT input_valid_a THEN
    channel_fault_a := channel_fault_a + 1;
END_IF;
cond_b := LimitHigh(raw_100_b, 120);
cond_b := cond_b AND quality_b;
cond_b := cond_b AND (NOT bypass_b);
input_valid_b := InputValid(raw_100_b, 0, 1000);
cond_b := cond_b AND input_valid_b;
IF NOT input_valid_b THEN
    channel_fault_b := channel_fault_b + 1;
END_IF;
cond_c := LimitHigh(raw_100_c, 120);
cond_c := cond_c AND quality_c;
cond_c := cond_c AND (NOT bypass_c);
input_valid_c := InputValid(raw_100_c, 0, 1000);
cond_c := cond_c AND input_valid_c;
IF NOT input_valid_c THEN
    channel_fault_c := channel_fault_c + 1;
END_IF;
cond_d := LimitHigh(raw_100_d, 120);
cond_d := cond_d AND quality_d;
cond_d := cond_d AND (NOT bypass_d);
input_valid_d := InputValid(raw_100_d, 0, 1000);
cond_d := cond_d AND input_valid_d;
IF NOT input_valid_d THEN
    channel_fault_d := channel_fault_d + 1;
END_IF;
vote_ok := TwoOfFour(cond_a, cond_b, cond_c, cond_d);
IF cond_a <> cond_b THEN
    diagnosis_count := diagnosis_count + 1;
END_IF;
IF cond_c <> cond_d THEN
    diagnosis_count := diagnosis_count + 1;
END_IF;
IF NOT vote_ok THEN
    diagnosis_count := diagnosis_count + 1;
END_IF;
latch_a_100 := RS_Next(vote_ok, train_a_reset, latch_a_100);
IF latch_a_100 AND (NOT train_a_inhibit) THEN
    mask_a_12 := mask_a_12 + 16;
    trip_a := 0 < 1;
    scram_a := 0 < 1;
    breaker_a := 0 > 1;
    si_a := 0 < 1;
    alarm_a := 0 < 1;
END_IF;
latch_b_100 := RS_Next(vote_ok, train_b_reset, latch_b_100);
IF latch_b_100 AND (NOT train_b_inhibit) THEN
    mask_b_12 := mask_b_12 + 16;
    trip_b := 0 < 1;
    scram_b := 0 < 1;
    breaker_b := 0 > 1;
    si_b := 0 < 1;
    alarm_b := 0 < 1;
END_IF;
IF (raw_100_a > 120) AND (NOT cond_a) THEN
    channel_fault_a := channel_fault_a + 1;
END_IF;
IF (raw_100_b > 120) AND (NOT cond_b) THEN
    channel_fault_b := channel_fault_b + 1;
END_IF;
IF (raw_100_c > 120) AND (NOT cond_c) THEN
    channel_fault_c := channel_fault_c + 1;
END_IF;
IF (raw_100_d > 120) AND (NOT cond_d) THEN
    channel_fault_d := channel_fault_d + 1;
END_IF;
IF vote_ok AND train_a_inhibit THEN
    diagnosis_count := diagnosis_count + 1;
END_IF;
IF vote_ok AND train_b_inhibit THEN
    diagnosis_count := diagnosis_count + 1;
END_IF;

cond_a := LimitHigh(raw_101_a, 121);
cond_a := cond_a AND quality_a;
cond_a := cond_a AND (NOT bypass_a);
input_valid_a := InputValid(raw_101_a, 0, 1000);
cond_a := cond_a AND input_valid_a;
IF NOT input_valid_a THEN
    channel_fault_a := channel_fault_a + 1;
END_IF;
cond_b := LimitHigh(raw_101_b, 121);
cond_b := cond_b AND quality_b;
cond_b := cond_b AND (NOT bypass_b);
input_valid_b := InputValid(raw_101_b, 0, 1000);
cond_b := cond_b AND input_valid_b;
IF NOT input_valid_b THEN
    channel_fault_b := channel_fault_b + 1;
END_IF;
cond_c := LimitHigh(raw_101_c, 121);
cond_c := cond_c AND quality_c;
cond_c := cond_c AND (NOT bypass_c);
input_valid_c := InputValid(raw_101_c, 0, 1000);
cond_c := cond_c AND input_valid_c;
IF NOT input_valid_c THEN
    channel_fault_c := channel_fault_c + 1;
END_IF;
cond_d := LimitHigh(raw_101_d, 121);
cond_d := cond_d AND quality_d;
cond_d := cond_d AND (NOT bypass_d);
input_valid_d := InputValid(raw_101_d, 0, 1000);
cond_d := cond_d AND input_valid_d;
IF NOT input_valid_d THEN
    channel_fault_d := channel_fault_d + 1;
END_IF;
vote_ok := TwoOfFour(cond_a, cond_b, cond_c, cond_d);
IF cond_a <> cond_b THEN
    diagnosis_count := diagnosis_count + 1;
END_IF;
IF cond_c <> cond_d THEN
    diagnosis_count := diagnosis_count + 1;
END_IF;
IF NOT vote_ok THEN
    diagnosis_count := diagnosis_count + 1;
END_IF;
latch_a_101 := RS_Next(vote_ok, train_a_reset, latch_a_101);
IF latch_a_101 AND (NOT train_a_inhibit) THEN
    mask_a_12 := mask_a_12 + 32;
    trip_a := 0 < 1;
    scram_a := 0 < 1;
    breaker_a := 0 > 1;
    ci_a := 0 < 1;
    alarm_a := 0 < 1;
END_IF;
latch_b_101 := RS_Next(vote_ok, train_b_reset, latch_b_101);
IF latch_b_101 AND (NOT train_b_inhibit) THEN
    mask_b_12 := mask_b_12 + 32;
    trip_b := 0 < 1;
    scram_b := 0 < 1;
    breaker_b := 0 > 1;
    ci_b := 0 < 1;
    alarm_b := 0 < 1;
END_IF;
IF (raw_101_a > 121) AND (NOT cond_a) THEN
    channel_fault_a := channel_fault_a + 1;
END_IF;
IF (raw_101_b > 121) AND (NOT cond_b) THEN
    channel_fault_b := channel_fault_b + 1;
END_IF;
IF (raw_101_c > 121) AND (NOT cond_c) THEN
    channel_fault_c := channel_fault_c + 1;
END_IF;
IF (raw_101_d > 121) AND (NOT cond_d) THEN
    channel_fault_d := channel_fault_d + 1;
END_IF;
IF vote_ok AND train_a_inhibit THEN
    diagnosis_count := diagnosis_count + 1;
END_IF;
IF vote_ok AND train_b_inhibit THEN
    diagnosis_count := diagnosis_count + 1;
END_IF;

cond_a := LimitHigh(raw_102_a, 122);
cond_a := cond_a AND quality_a;
cond_a := cond_a AND (NOT bypass_a);
input_valid_a := InputValid(raw_102_a, 0, 1000);
cond_a := cond_a AND input_valid_a;
IF NOT input_valid_a THEN
    channel_fault_a := channel_fault_a + 1;
END_IF;
cond_b := LimitHigh(raw_102_b, 122);
cond_b := cond_b AND quality_b;
cond_b := cond_b AND (NOT bypass_b);
input_valid_b := InputValid(raw_102_b, 0, 1000);
cond_b := cond_b AND input_valid_b;
IF NOT input_valid_b THEN
    channel_fault_b := channel_fault_b + 1;
END_IF;
cond_c := LimitHigh(raw_102_c, 122);
cond_c := cond_c AND quality_c;
cond_c := cond_c AND (NOT bypass_c);
input_valid_c := InputValid(raw_102_c, 0, 1000);
cond_c := cond_c AND input_valid_c;
IF NOT input_valid_c THEN
    channel_fault_c := channel_fault_c + 1;
END_IF;
cond_d := LimitHigh(raw_102_d, 122);
cond_d := cond_d AND quality_d;
cond_d := cond_d AND (NOT bypass_d);
input_valid_d := InputValid(raw_102_d, 0, 1000);
cond_d := cond_d AND input_valid_d;
IF NOT input_valid_d THEN
    channel_fault_d := channel_fault_d + 1;
END_IF;
vote_ok := TwoOfFour(cond_a, cond_b, cond_c, cond_d);
IF cond_a <> cond_b THEN
    diagnosis_count := diagnosis_count + 1;
END_IF;
IF cond_c <> cond_d THEN
    diagnosis_count := diagnosis_count + 1;
END_IF;
IF NOT vote_ok THEN
    diagnosis_count := diagnosis_count + 1;
END_IF;
latch_a_102 := RS_Next(vote_ok, train_a_reset, latch_a_102);
IF latch_a_102 AND (NOT train_a_inhibit) THEN
    mask_a_12 := mask_a_12 + 64;
    trip_a := 0 < 1;
    scram_a := 0 < 1;
    breaker_a := 0 > 1;
    mfw_a := 0 < 1;
    alarm_a := 0 < 1;
END_IF;
latch_b_102 := RS_Next(vote_ok, train_b_reset, latch_b_102);
IF latch_b_102 AND (NOT train_b_inhibit) THEN
    mask_b_12 := mask_b_12 + 64;
    trip_b := 0 < 1;
    scram_b := 0 < 1;
    breaker_b := 0 > 1;
    mfw_b := 0 < 1;
    alarm_b := 0 < 1;
END_IF;
IF (raw_102_a > 122) AND (NOT cond_a) THEN
    channel_fault_a := channel_fault_a + 1;
END_IF;
IF (raw_102_b > 122) AND (NOT cond_b) THEN
    channel_fault_b := channel_fault_b + 1;
END_IF;
IF (raw_102_c > 122) AND (NOT cond_c) THEN
    channel_fault_c := channel_fault_c + 1;
END_IF;
IF (raw_102_d > 122) AND (NOT cond_d) THEN
    channel_fault_d := channel_fault_d + 1;
END_IF;
IF vote_ok AND train_a_inhibit THEN
    diagnosis_count := diagnosis_count + 1;
END_IF;
IF vote_ok AND train_b_inhibit THEN
    diagnosis_count := diagnosis_count + 1;
END_IF;

cond_a := LimitHigh(raw_103_a, 123);
cond_a := cond_a AND quality_a;
cond_a := cond_a AND (NOT bypass_a);
input_valid_a := InputValid(raw_103_a, 0, 1000);
cond_a := cond_a AND input_valid_a;
IF NOT input_valid_a THEN
    channel_fault_a := channel_fault_a + 1;
END_IF;
cond_b := LimitHigh(raw_103_b, 123);
cond_b := cond_b AND quality_b;
cond_b := cond_b AND (NOT bypass_b);
input_valid_b := InputValid(raw_103_b, 0, 1000);
cond_b := cond_b AND input_valid_b;
IF NOT input_valid_b THEN
    channel_fault_b := channel_fault_b + 1;
END_IF;
cond_c := LimitHigh(raw_103_c, 123);
cond_c := cond_c AND quality_c;
cond_c := cond_c AND (NOT bypass_c);
input_valid_c := InputValid(raw_103_c, 0, 1000);
cond_c := cond_c AND input_valid_c;
IF NOT input_valid_c THEN
    channel_fault_c := channel_fault_c + 1;
END_IF;
cond_d := LimitHigh(raw_103_d, 123);
cond_d := cond_d AND quality_d;
cond_d := cond_d AND (NOT bypass_d);
input_valid_d := InputValid(raw_103_d, 0, 1000);
cond_d := cond_d AND input_valid_d;
IF NOT input_valid_d THEN
    channel_fault_d := channel_fault_d + 1;
END_IF;
vote_ok := TwoOfFour(cond_a, cond_b, cond_c, cond_d);
IF cond_a <> cond_b THEN
    diagnosis_count := diagnosis_count + 1;
END_IF;
IF cond_c <> cond_d THEN
    diagnosis_count := diagnosis_count + 1;
END_IF;
IF NOT vote_ok THEN
    diagnosis_count := diagnosis_count + 1;
END_IF;
latch_a_103 := RS_Next(vote_ok, train_a_reset, latch_a_103);
IF latch_a_103 AND (NOT train_a_inhibit) THEN
    mask_a_12 := mask_a_12 + 128;
    trip_a := 0 < 1;
    scram_a := 0 < 1;
    breaker_a := 0 > 1;
    afw_a := 0 < 1;
    alarm_a := 0 < 1;
END_IF;
latch_b_103 := RS_Next(vote_ok, train_b_reset, latch_b_103);
IF latch_b_103 AND (NOT train_b_inhibit) THEN
    mask_b_12 := mask_b_12 + 128;
    trip_b := 0 < 1;
    scram_b := 0 < 1;
    breaker_b := 0 > 1;
    afw_b := 0 < 1;
    alarm_b := 0 < 1;
END_IF;
IF (raw_103_a > 123) AND (NOT cond_a) THEN
    channel_fault_a := channel_fault_a + 1;
END_IF;
IF (raw_103_b > 123) AND (NOT cond_b) THEN
    channel_fault_b := channel_fault_b + 1;
END_IF;
IF (raw_103_c > 123) AND (NOT cond_c) THEN
    channel_fault_c := channel_fault_c + 1;
END_IF;
IF (raw_103_d > 123) AND (NOT cond_d) THEN
    channel_fault_d := channel_fault_d + 1;
END_IF;
IF vote_ok AND train_a_inhibit THEN
    diagnosis_count := diagnosis_count + 1;
END_IF;
IF vote_ok AND train_b_inhibit THEN
    diagnosis_count := diagnosis_count + 1;
END_IF;

cond_a := LimitHigh(raw_104_a, 124);
cond_a := cond_a AND quality_a;
cond_a := cond_a AND (NOT bypass_a);
input_valid_a := InputValid(raw_104_a, 0, 1000);
cond_a := cond_a AND input_valid_a;
IF NOT input_valid_a THEN
    channel_fault_a := channel_fault_a + 1;
END_IF;
cond_b := LimitHigh(raw_104_b, 124);
cond_b := cond_b AND quality_b;
cond_b := cond_b AND (NOT bypass_b);
input_valid_b := InputValid(raw_104_b, 0, 1000);
cond_b := cond_b AND input_valid_b;
IF NOT input_valid_b THEN
    channel_fault_b := channel_fault_b + 1;
END_IF;
cond_c := LimitHigh(raw_104_c, 124);
cond_c := cond_c AND quality_c;
cond_c := cond_c AND (NOT bypass_c);
input_valid_c := InputValid(raw_104_c, 0, 1000);
cond_c := cond_c AND input_valid_c;
IF NOT input_valid_c THEN
    channel_fault_c := channel_fault_c + 1;
END_IF;
cond_d := LimitHigh(raw_104_d, 124);
cond_d := cond_d AND quality_d;
cond_d := cond_d AND (NOT bypass_d);
input_valid_d := InputValid(raw_104_d, 0, 1000);
cond_d := cond_d AND input_valid_d;
IF NOT input_valid_d THEN
    channel_fault_d := channel_fault_d + 1;
END_IF;
vote_ok := TwoOfFour(cond_a, cond_b, cond_c, cond_d);
IF cond_a <> cond_b THEN
    diagnosis_count := diagnosis_count + 1;
END_IF;
IF cond_c <> cond_d THEN
    diagnosis_count := diagnosis_count + 1;
END_IF;
IF NOT vote_ok THEN
    diagnosis_count := diagnosis_count + 1;
END_IF;
latch_a_104 := RS_Next(vote_ok, train_a_reset, latch_a_104);
IF latch_a_104 AND (NOT train_a_inhibit) THEN
    mask_a_13 := mask_a_13 + 1;
    trip_a := 0 < 1;
    scram_a := 0 < 1;
    breaker_a := 0 > 1;
    si_a := 0 < 1;
    alarm_a := 0 < 1;
END_IF;
latch_b_104 := RS_Next(vote_ok, train_b_reset, latch_b_104);
IF latch_b_104 AND (NOT train_b_inhibit) THEN
    mask_b_13 := mask_b_13 + 1;
    trip_b := 0 < 1;
    scram_b := 0 < 1;
    breaker_b := 0 > 1;
    si_b := 0 < 1;
    alarm_b := 0 < 1;
END_IF;
IF (raw_104_a > 124) AND (NOT cond_a) THEN
    channel_fault_a := channel_fault_a + 1;
END_IF;
IF (raw_104_b > 124) AND (NOT cond_b) THEN
    channel_fault_b := channel_fault_b + 1;
END_IF;
IF (raw_104_c > 124) AND (NOT cond_c) THEN
    channel_fault_c := channel_fault_c + 1;
END_IF;
IF (raw_104_d > 124) AND (NOT cond_d) THEN
    channel_fault_d := channel_fault_d + 1;
END_IF;
IF vote_ok AND train_a_inhibit THEN
    diagnosis_count := diagnosis_count + 1;
END_IF;
IF vote_ok AND train_b_inhibit THEN
    diagnosis_count := diagnosis_count + 1;
END_IF;

cond_a := LimitHigh(raw_105_a, 125);
cond_a := cond_a AND quality_a;
cond_a := cond_a AND (NOT bypass_a);
input_valid_a := InputValid(raw_105_a, 0, 1000);
cond_a := cond_a AND input_valid_a;
IF NOT input_valid_a THEN
    channel_fault_a := channel_fault_a + 1;
END_IF;
cond_b := LimitHigh(raw_105_b, 125);
cond_b := cond_b AND quality_b;
cond_b := cond_b AND (NOT bypass_b);
input_valid_b := InputValid(raw_105_b, 0, 1000);
cond_b := cond_b AND input_valid_b;
IF NOT input_valid_b THEN
    channel_fault_b := channel_fault_b + 1;
END_IF;
cond_c := LimitHigh(raw_105_c, 125);
cond_c := cond_c AND quality_c;
cond_c := cond_c AND (NOT bypass_c);
input_valid_c := InputValid(raw_105_c, 0, 1000);
cond_c := cond_c AND input_valid_c;
IF NOT input_valid_c THEN
    channel_fault_c := channel_fault_c + 1;
END_IF;
cond_d := LimitHigh(raw_105_d, 125);
cond_d := cond_d AND quality_d;
cond_d := cond_d AND (NOT bypass_d);
input_valid_d := InputValid(raw_105_d, 0, 1000);
cond_d := cond_d AND input_valid_d;
IF NOT input_valid_d THEN
    channel_fault_d := channel_fault_d + 1;
END_IF;
vote_ok := TwoOfFour(cond_a, cond_b, cond_c, cond_d);
IF cond_a <> cond_b THEN
    diagnosis_count := diagnosis_count + 1;
END_IF;
IF cond_c <> cond_d THEN
    diagnosis_count := diagnosis_count + 1;
END_IF;
IF NOT vote_ok THEN
    diagnosis_count := diagnosis_count + 1;
END_IF;
latch_a_105 := RS_Next(vote_ok, train_a_reset, latch_a_105);
IF latch_a_105 AND (NOT train_a_inhibit) THEN
    mask_a_13 := mask_a_13 + 2;
    trip_a := 0 < 1;
    scram_a := 0 < 1;
    breaker_a := 0 > 1;
    ci_a := 0 < 1;
    alarm_a := 0 < 1;
END_IF;
latch_b_105 := RS_Next(vote_ok, train_b_reset, latch_b_105);
IF latch_b_105 AND (NOT train_b_inhibit) THEN
    mask_b_13 := mask_b_13 + 2;
    trip_b := 0 < 1;
    scram_b := 0 < 1;
    breaker_b := 0 > 1;
    ci_b := 0 < 1;
    alarm_b := 0 < 1;
END_IF;
IF (raw_105_a > 125) AND (NOT cond_a) THEN
    channel_fault_a := channel_fault_a + 1;
END_IF;
IF (raw_105_b > 125) AND (NOT cond_b) THEN
    channel_fault_b := channel_fault_b + 1;
END_IF;
IF (raw_105_c > 125) AND (NOT cond_c) THEN
    channel_fault_c := channel_fault_c + 1;
END_IF;
IF (raw_105_d > 125) AND (NOT cond_d) THEN
    channel_fault_d := channel_fault_d + 1;
END_IF;
IF vote_ok AND train_a_inhibit THEN
    diagnosis_count := diagnosis_count + 1;
END_IF;
IF vote_ok AND train_b_inhibit THEN
    diagnosis_count := diagnosis_count + 1;
END_IF;

cond_a := LimitHigh(raw_106_a, 126);
cond_a := cond_a AND quality_a;
cond_a := cond_a AND (NOT bypass_a);
input_valid_a := InputValid(raw_106_a, 0, 1000);
cond_a := cond_a AND input_valid_a;
IF NOT input_valid_a THEN
    channel_fault_a := channel_fault_a + 1;
END_IF;
cond_b := LimitHigh(raw_106_b, 126);
cond_b := cond_b AND quality_b;
cond_b := cond_b AND (NOT bypass_b);
input_valid_b := InputValid(raw_106_b, 0, 1000);
cond_b := cond_b AND input_valid_b;
IF NOT input_valid_b THEN
    channel_fault_b := channel_fault_b + 1;
END_IF;
cond_c := LimitHigh(raw_106_c, 126);
cond_c := cond_c AND quality_c;
cond_c := cond_c AND (NOT bypass_c);
input_valid_c := InputValid(raw_106_c, 0, 1000);
cond_c := cond_c AND input_valid_c;
IF NOT input_valid_c THEN
    channel_fault_c := channel_fault_c + 1;
END_IF;
cond_d := LimitHigh(raw_106_d, 126);
cond_d := cond_d AND quality_d;
cond_d := cond_d AND (NOT bypass_d);
input_valid_d := InputValid(raw_106_d, 0, 1000);
cond_d := cond_d AND input_valid_d;
IF NOT input_valid_d THEN
    channel_fault_d := channel_fault_d + 1;
END_IF;
vote_ok := TwoOfFour(cond_a, cond_b, cond_c, cond_d);
IF cond_a <> cond_b THEN
    diagnosis_count := diagnosis_count + 1;
END_IF;
IF cond_c <> cond_d THEN
    diagnosis_count := diagnosis_count + 1;
END_IF;
IF NOT vote_ok THEN
    diagnosis_count := diagnosis_count + 1;
END_IF;
latch_a_106 := RS_Next(vote_ok, train_a_reset, latch_a_106);
IF latch_a_106 AND (NOT train_a_inhibit) THEN
    mask_a_13 := mask_a_13 + 4;
    trip_a := 0 < 1;
    scram_a := 0 < 1;
    breaker_a := 0 > 1;
    mfw_a := 0 < 1;
    alarm_a := 0 < 1;
END_IF;
latch_b_106 := RS_Next(vote_ok, train_b_reset, latch_b_106);
IF latch_b_106 AND (NOT train_b_inhibit) THEN
    mask_b_13 := mask_b_13 + 4;
    trip_b := 0 < 1;
    scram_b := 0 < 1;
    breaker_b := 0 > 1;
    mfw_b := 0 < 1;
    alarm_b := 0 < 1;
END_IF;
IF (raw_106_a > 126) AND (NOT cond_a) THEN
    channel_fault_a := channel_fault_a + 1;
END_IF;
IF (raw_106_b > 126) AND (NOT cond_b) THEN
    channel_fault_b := channel_fault_b + 1;
END_IF;
IF (raw_106_c > 126) AND (NOT cond_c) THEN
    channel_fault_c := channel_fault_c + 1;
END_IF;
IF (raw_106_d > 126) AND (NOT cond_d) THEN
    channel_fault_d := channel_fault_d + 1;
END_IF;
IF vote_ok AND train_a_inhibit THEN
    diagnosis_count := diagnosis_count + 1;
END_IF;
IF vote_ok AND train_b_inhibit THEN
    diagnosis_count := diagnosis_count + 1;
END_IF;

cond_a := LimitHigh(raw_107_a, 127);
cond_a := cond_a AND quality_a;
cond_a := cond_a AND (NOT bypass_a);
input_valid_a := InputValid(raw_107_a, 0, 1000);
cond_a := cond_a AND input_valid_a;
IF NOT input_valid_a THEN
    channel_fault_a := channel_fault_a + 1;
END_IF;
cond_b := LimitHigh(raw_107_b, 127);
cond_b := cond_b AND quality_b;
cond_b := cond_b AND (NOT bypass_b);
input_valid_b := InputValid(raw_107_b, 0, 1000);
cond_b := cond_b AND input_valid_b;
IF NOT input_valid_b THEN
    channel_fault_b := channel_fault_b + 1;
END_IF;
cond_c := LimitHigh(raw_107_c, 127);
cond_c := cond_c AND quality_c;
cond_c := cond_c AND (NOT bypass_c);
input_valid_c := InputValid(raw_107_c, 0, 1000);
cond_c := cond_c AND input_valid_c;
IF NOT input_valid_c THEN
    channel_fault_c := channel_fault_c + 1;
END_IF;
cond_d := LimitHigh(raw_107_d, 127);
cond_d := cond_d AND quality_d;
cond_d := cond_d AND (NOT bypass_d);
input_valid_d := InputValid(raw_107_d, 0, 1000);
cond_d := cond_d AND input_valid_d;
IF NOT input_valid_d THEN
    channel_fault_d := channel_fault_d + 1;
END_IF;
vote_ok := TwoOfFour(cond_a, cond_b, cond_c, cond_d);
IF cond_a <> cond_b THEN
    diagnosis_count := diagnosis_count + 1;
END_IF;
IF cond_c <> cond_d THEN
    diagnosis_count := diagnosis_count + 1;
END_IF;
IF NOT vote_ok THEN
    diagnosis_count := diagnosis_count + 1;
END_IF;
latch_a_107 := RS_Next(vote_ok, train_a_reset, latch_a_107);
IF latch_a_107 AND (NOT train_a_inhibit) THEN
    mask_a_13 := mask_a_13 + 8;
    trip_a := 0 < 1;
    scram_a := 0 < 1;
    breaker_a := 0 > 1;
    afw_a := 0 < 1;
    alarm_a := 0 < 1;
END_IF;
latch_b_107 := RS_Next(vote_ok, train_b_reset, latch_b_107);
IF latch_b_107 AND (NOT train_b_inhibit) THEN
    mask_b_13 := mask_b_13 + 8;
    trip_b := 0 < 1;
    scram_b := 0 < 1;
    breaker_b := 0 > 1;
    afw_b := 0 < 1;
    alarm_b := 0 < 1;
END_IF;
IF (raw_107_a > 127) AND (NOT cond_a) THEN
    channel_fault_a := channel_fault_a + 1;
END_IF;
IF (raw_107_b > 127) AND (NOT cond_b) THEN
    channel_fault_b := channel_fault_b + 1;
END_IF;
IF (raw_107_c > 127) AND (NOT cond_c) THEN
    channel_fault_c := channel_fault_c + 1;
END_IF;
IF (raw_107_d > 127) AND (NOT cond_d) THEN
    channel_fault_d := channel_fault_d + 1;
END_IF;
IF vote_ok AND train_a_inhibit THEN
    diagnosis_count := diagnosis_count + 1;
END_IF;
IF vote_ok AND train_b_inhibit THEN
    diagnosis_count := diagnosis_count + 1;
END_IF;

cond_a := LimitHigh(raw_108_a, 128);
cond_a := cond_a AND quality_a;
cond_a := cond_a AND (NOT bypass_a);
input_valid_a := InputValid(raw_108_a, 0, 1000);
cond_a := cond_a AND input_valid_a;
IF NOT input_valid_a THEN
    channel_fault_a := channel_fault_a + 1;
END_IF;
cond_b := LimitHigh(raw_108_b, 128);
cond_b := cond_b AND quality_b;
cond_b := cond_b AND (NOT bypass_b);
input_valid_b := InputValid(raw_108_b, 0, 1000);
cond_b := cond_b AND input_valid_b;
IF NOT input_valid_b THEN
    channel_fault_b := channel_fault_b + 1;
END_IF;
cond_c := LimitHigh(raw_108_c, 128);
cond_c := cond_c AND quality_c;
cond_c := cond_c AND (NOT bypass_c);
input_valid_c := InputValid(raw_108_c, 0, 1000);
cond_c := cond_c AND input_valid_c;
IF NOT input_valid_c THEN
    channel_fault_c := channel_fault_c + 1;
END_IF;
cond_d := LimitHigh(raw_108_d, 128);
cond_d := cond_d AND quality_d;
cond_d := cond_d AND (NOT bypass_d);
input_valid_d := InputValid(raw_108_d, 0, 1000);
cond_d := cond_d AND input_valid_d;
IF NOT input_valid_d THEN
    channel_fault_d := channel_fault_d + 1;
END_IF;
vote_ok := TwoOfFour(cond_a, cond_b, cond_c, cond_d);
IF cond_a <> cond_b THEN
    diagnosis_count := diagnosis_count + 1;
END_IF;
IF cond_c <> cond_d THEN
    diagnosis_count := diagnosis_count + 1;
END_IF;
IF NOT vote_ok THEN
    diagnosis_count := diagnosis_count + 1;
END_IF;
latch_a_108 := RS_Next(vote_ok, train_a_reset, latch_a_108);
IF latch_a_108 AND (NOT train_a_inhibit) THEN
    mask_a_13 := mask_a_13 + 16;
    trip_a := 0 < 1;
    scram_a := 0 < 1;
    breaker_a := 0 > 1;
    si_a := 0 < 1;
    alarm_a := 0 < 1;
END_IF;
latch_b_108 := RS_Next(vote_ok, train_b_reset, latch_b_108);
IF latch_b_108 AND (NOT train_b_inhibit) THEN
    mask_b_13 := mask_b_13 + 16;
    trip_b := 0 < 1;
    scram_b := 0 < 1;
    breaker_b := 0 > 1;
    si_b := 0 < 1;
    alarm_b := 0 < 1;
END_IF;
IF (raw_108_a > 128) AND (NOT cond_a) THEN
    channel_fault_a := channel_fault_a + 1;
END_IF;
IF (raw_108_b > 128) AND (NOT cond_b) THEN
    channel_fault_b := channel_fault_b + 1;
END_IF;
IF (raw_108_c > 128) AND (NOT cond_c) THEN
    channel_fault_c := channel_fault_c + 1;
END_IF;
IF (raw_108_d > 128) AND (NOT cond_d) THEN
    channel_fault_d := channel_fault_d + 1;
END_IF;
IF vote_ok AND train_a_inhibit THEN
    diagnosis_count := diagnosis_count + 1;
END_IF;
IF vote_ok AND train_b_inhibit THEN
    diagnosis_count := diagnosis_count + 1;
END_IF;

cond_a := LimitHigh(raw_109_a, 129);
cond_a := cond_a AND quality_a;
cond_a := cond_a AND (NOT bypass_a);
input_valid_a := InputValid(raw_109_a, 0, 1000);
cond_a := cond_a AND input_valid_a;
IF NOT input_valid_a THEN
    channel_fault_a := channel_fault_a + 1;
END_IF;
cond_b := LimitHigh(raw_109_b, 129);
cond_b := cond_b AND quality_b;
cond_b := cond_b AND (NOT bypass_b);
input_valid_b := InputValid(raw_109_b, 0, 1000);
cond_b := cond_b AND input_valid_b;
IF NOT input_valid_b THEN
    channel_fault_b := channel_fault_b + 1;
END_IF;
cond_c := LimitHigh(raw_109_c, 129);
cond_c := cond_c AND quality_c;
cond_c := cond_c AND (NOT bypass_c);
input_valid_c := InputValid(raw_109_c, 0, 1000);
cond_c := cond_c AND input_valid_c;
IF NOT input_valid_c THEN
    channel_fault_c := channel_fault_c + 1;
END_IF;
cond_d := LimitHigh(raw_109_d, 129);
cond_d := cond_d AND quality_d;
cond_d := cond_d AND (NOT bypass_d);
input_valid_d := InputValid(raw_109_d, 0, 1000);
cond_d := cond_d AND input_valid_d;
IF NOT input_valid_d THEN
    channel_fault_d := channel_fault_d + 1;
END_IF;
vote_ok := TwoOfFour(cond_a, cond_b, cond_c, cond_d);
IF cond_a <> cond_b THEN
    diagnosis_count := diagnosis_count + 1;
END_IF;
IF cond_c <> cond_d THEN
    diagnosis_count := diagnosis_count + 1;
END_IF;
IF NOT vote_ok THEN
    diagnosis_count := diagnosis_count + 1;
END_IF;
latch_a_109 := RS_Next(vote_ok, train_a_reset, latch_a_109);
IF latch_a_109 AND (NOT train_a_inhibit) THEN
    mask_a_13 := mask_a_13 + 32;
    trip_a := 0 < 1;
    scram_a := 0 < 1;
    breaker_a := 0 > 1;
    ci_a := 0 < 1;
    alarm_a := 0 < 1;
END_IF;
latch_b_109 := RS_Next(vote_ok, train_b_reset, latch_b_109);
IF latch_b_109 AND (NOT train_b_inhibit) THEN
    mask_b_13 := mask_b_13 + 32;
    trip_b := 0 < 1;
    scram_b := 0 < 1;
    breaker_b := 0 > 1;
    ci_b := 0 < 1;
    alarm_b := 0 < 1;
END_IF;
IF (raw_109_a > 129) AND (NOT cond_a) THEN
    channel_fault_a := channel_fault_a + 1;
END_IF;
IF (raw_109_b > 129) AND (NOT cond_b) THEN
    channel_fault_b := channel_fault_b + 1;
END_IF;
IF (raw_109_c > 129) AND (NOT cond_c) THEN
    channel_fault_c := channel_fault_c + 1;
END_IF;
IF (raw_109_d > 129) AND (NOT cond_d) THEN
    channel_fault_d := channel_fault_d + 1;
END_IF;
IF vote_ok AND train_a_inhibit THEN
    diagnosis_count := diagnosis_count + 1;
END_IF;
IF vote_ok AND train_b_inhibit THEN
    diagnosis_count := diagnosis_count + 1;
END_IF;
